_articlenumberRegex	:= '';
_serialnumberRegex	:= '';
_traceID						:= DINT#0;
_activeCheckFQDN		:= FALSE;
_allowedFQDN				:= '';

_previousProcesses.Clear();
END_METHOD

METHOD PUBLIC CopyFrom : BOOL
VAR_INPUT
	IN	: KOSTAL_AF2024_Core_System.I_Interface;
END_VAR

VAR
	_IN		: I_T_ProcessConfig;
//	_udi	: UDINT;
//	_p		: POINTER TO T_PreviousProcess;
//	_resp	: KOSTAL_AF2024_Core_functionResponse.T_functionResponse;
END_VAR

IF NOT SUPER^.CopyFrom(IN) 												THEN RETURN;	END_IF
IF NOT __QUERYINTERFACE(IN, _IN) OR_ELSE _IN = 0 	THEN RETURN;	END_IF

_serialnumberRegex	:= _IN.serialnumberRegex;
_articlenumberRegex	:= _IN.articlenumberRegex;
_traceId						:= _IN.traceId;
_activeCheckFQDN		:= _IN.activeCheckFQDN;
_allowedFQDN				:= _IN.allowedFQDN;

_previousProcesses.CopyFrom(_IN.PreviousProcesses);

CopyFrom:= TRUE;

//FOR _udi:= 1 TO _IN.PreviousProcesses.NumberOfObjects DO

//	IF NOT _previousProcesses.AddObject() THEN RETURN;	END_IF

//	_p:= 	_previousProcesses.Get_P(_previousProcesses.NumberOfObjects, _resp);

//	IF (NOT _resp.success) OR (_p = 0 ) THEN RETURN;	END_IF
	
//	_p^.CopyFrom(IN.IPreviousProcesses.Get_I(_udi, _resp));
		
//END_FOR
END_METHOD

PROPERTY PUBLIC PreviousProcesses : I_ListOfPreviousProcess
GET

PreviousProcesses:= _previousProcesses;
END_GET
END_PROPERTY

PROPERTY PUBLIC PreviousProcesses_Owner : I_ListOfPreviousProcess_Owner
GET

PreviousProcesses_Owner := _previousProcesses;
END_GET
END_PROPERTY

PROPERTY PUBLIC serialnumberRegex : KOSTAL_AF2024_Core_Settings.T_MaxString_UTF8
GET

serialnumberRegex:= _serialnumberRegex;
END_GET
SET

_serialnumberRegex:= serialnumberRegex;
END_SET
END_PROPERTY

PROPERTY PUBLIC traceID : DINT
GET

traceID:= _traceID;
END_GET
SET

_traceID:= traceID;
END_SET
END_PROPERTY

END_FUNCTION_BLOCK

// 3_DUT/SingleProcess/ListOf/FB_ListOfSingleProcess
FUNCTION_BLOCK FB_ListOfSingleProcess  EXTENDS KOSTAL_AF2024_Core_ListOf._FB_Object_Base IMPLEMENTS I_ListOfSingleProcess, I_ListOfSingleProcess_CopyFrom, I_ListOfSingleProcess_Owner

VAR
	_Dummy	: T_SingleProcess;
END_VAR

(*
	Returns the typed interface in the reference variable.
	In the event of an error, the return value becomes FALSE and the interface refers to the {_Dummy}.
*)
METHOD PROTECTED _get_I : I_T_SingleProcess

VAR_INPUT
	Member		: KOSTAL_AF2024_Core_System.I_Interface;
	rValid		: REFERENCE TO BOOL;
	Response	: KOSTAL_AF2024_Core_functionResponse.I_T_functionResponse_Owner;
END_VAR

VAR
	_iObj			: I_T_SingleProcess;
END_VAR
//preset
_get_I:= _Dummy;
IF __ISVALIDREF(rValid)	THEN	rValid:= FALSE;	END_IF	

IF NOT _verifyMember(Member, Response)	THEN RETURN;	END_IF

//return dummy if no valid DUT is found
IF NOT __QUERYINTERFACE(Member, _iObj) OR_ELSE (_iObj = 0)	THEN		
	_setResultFail(Response, "__QueryInterface failed - return Dummy");	RETURN;	
END_IF

IF __ISVALIDREF(rValid)	THEN	rValid:= TRUE;	END_IF	
_setResultPass(Response, "Successful");

_get_I:= _iObj;
END_METHOD

(*
	Returns the typed owner interface in the reference variable.
	In the event of an error, the return value becomes FALSE and the interface refers to the {_Dummy}.
*)
METHOD PROTECTED _get_I_Owner : I_T_SingleProcess_Owner

VAR_INPUT
	Member		: KOSTAL_AF2024_Core_System.I_Interface;
	rValid		: REFERENCE TO BOOL;
	Response	: KOSTAL_AF2024_Core_functionResponse.I_T_functionResponse_Owner;
END_VAR

VAR
	_iObj			: I_T_SingleProcess_Owner;
END_VAR
//preset
_get_I_Owner:= _Dummy;

IF 		__ISVALIDREF(rValid)	THEN	rValid:= FALSE;	END_IF	

IF NOT _verifyMember(Member, Response)	THEN RETURN;	END_IF

//return dummy if no valid DUT is found
IF NOT __QUERYINTERFACE(Member, _iObj) OR_ELSE (_iObj = 0)	THEN	
	_setResultFail(Response, "__QueryInterface failed - return Dummy");	RETURN;	
END_IF

IF __ISVALIDREF(rValid)	THEN	rValid:= TRUE;	END_IF
_setResultPass(Response, "Successful");
_get_I_Owner:= _iObj;
END_METHOD

(*
	Cleans the custom class {FB_DUT} and removes it from memory.
*)
METHOD PROTECTED  _removePayLoad : BOOL
VAR_INPUT
	Member	: KOSTAL_AF2024_Core_System.I_Interface;
	Result	: KOSTAL_AF2024_Core_functionResponse.I_T_functionResponse_Owner;
END_VAR

VAR
	_iObj			: I_T_SingleProcess_Owner;
	_pFB_DUT	:	POINTER TO T_SingleProcess;
	_Success	: BOOL;
END_VAR


IF NOT SUPER^._removePayload(Member, Result)	THEN RETURN;	END_IF

_Success:= __QUERYINTERFACE(Member, _iObj);

IF NOT _Success	THEN	RETURN;	END_IF
IF _iObj = 0		THEN	RETURN;	END_IF

_iObj.Clear();

_Success  := __QUERYPOINTER(_iObj, _pFB_DUT);

IF NOT _Success	THEN	RETURN;	END_IF
IF _pFB_DUT = 0	THEN	RETURN;	END_IF

__DELETE(_pFB_DUT);
END_METHOD

(*
	Overload the method from the base class to verify the custom interface. 
	The local method {_get_I_Owner()} is used for this.
*)
METHOD PROTECTED _verifyMember : BOOL

VAR_INPUT
	Member	: KOSTAL_AF2024_Core_System.I_Interface;
	Result	: KOSTAL_AF2024_Core_functionResponse.I_T_functionResponse_Owner;
END_VAR

VAR
	_pObj	: POINTER TO T_SingleProcess;
	_Success: BOOL;
END_VAR

IF NOT SUPER^._verifyMember(Member, Result)	THEN RETURN;	END_IF

_Success:= __QUERYPOINTER(Member, _pObj);

//return dummy if no valid Pointer to DUT is found
IF NOT _Success OR_ELSE (_pObj = 0)	THEN	_setResultFail(Result, "__QueryPointer failed");	RETURN; END_IF

_verifyMember:= TRUE;
END_METHOD

(*
	Add a new instance of FB_Dut and copy content from [IN] to the new instance
*)
METHOD PUBLIC Add_DUT : BOOL
VAR_INPUT
	IN				: KOSTAL_AF2024_Core_System.I_Interface;
	Response	: KOSTAL_AF2024_Core_functionResponse.I_T_functionResponse_Owner;
END_VAR

VAR
	_IN1	: I_T_SingleProcess;
	_IN2	: I_T_SingleProcess_Owner;
	_pDUT	: POINTER TO T_SingleProcess;
END_VAR

IF IN = 0 THEN	RETURN;	END_IF


IF __QUERYINTERFACE(IN, _IN1) AND_THEN (_IN1 <> 0)	THEN


	_pDUT:= __NEW(T_SingleProcess);
	
	IF _pDUT = 0 THEN	_setResultFail(Response, "cannot create new object"); RETURN; END_IF
	
	_pDUT^.CopyFrom(_IN1);
	
	Add_DUT:= _addMember(_pDUT^, Response);


ELSIF __QUERYINTERFACE(IN, _IN2) AND_THEN (_IN2 <> 0)	THEN


	_pDUT:= __NEW(T_SingleProcess);
	
	IF _pDUT = 0 THEN	_setResultFail(Response, "cannot create new object"); RETURN; END_IF
	
	_pDUT^.CopyFrom(_IN2);
	
	Add_DUT:= _addMember(_pDUT^, Response);


END_IF
END_METHOD

(*
	Makes the protected method public.
*)
METHOD Clear

_clear();
END_METHOD

(*
	Copies the contents of another list {IN} into its own memory.
*)
METHOD PUBLIC CopyFrom
VAR_INPUT
	IN	: KOSTAL_AF2024_Core_System.I_Interface;
END_VAR

VAR
	_udi	: UDINT;

	_IN		: I_ListOfSingleProcess;
	_IN_O	: I_ListOfSingleProcess_Owner;

END_VAR

IF IN = 0 THEN RETURN;	END_IF

IF __QUERYINTERFACE(IN, _IN_O) AND_THEN _IN_O <> 0	THEN

	_clear();
	
	FOR _udi:= 1 TO _IN_O.NumberOfMember DO
		Add_DUT(_IN_O.Get_I_Owner(_udi, 0, 0), 0);
	END_FOR
	
ELSIF __QUERYINTERFACE(IN, _IN) AND_THEN _IN <> 0	THEN	

	_clear();
	
	FOR _udi:= 1 TO _IN.NumberOfMember DO
		Add_DUT(_IN.Get_I(_udi, 0, 0), 0);
	END_FOR

END_IF
END_METHOD

(*
	Copies the own content into another list created at the parameter {IN}.
*)
METHOD PUBLIC CopyTo
VAR_INPUT
	IN	: KOSTAL_AF2024_Core_System.I_Interface;
END_VAR

VAR
	_IN	: I_ListOfSingleProcess_CopyFrom;
END_VAR

IF (IN = 0) OR_ELSE NOT __QUERYINTERFACE(IN, _IN) OR_ELSE (_IN = 0) THEN	RETURN;	END_IF

_IN.CopyFrom(THIS^);
END_METHOD

(*
	Deletes the class specified with the {Number} from the list.
*)
METHOD PUBLIC Delete_DUT : BOOL
VAR_INPUT
	Number		: UDINT;	//Number of DUT in List
	Response	: KOSTAL_AF2024_Core_functionResponse.I_T_functionResponse_Owner;
END_VAR

VAR
	//_response	: KOSTAL_AF2024_Core_functionResponse.T_functionResponse;
	_Success	: BOOL;
	_Member		: KOSTAL_AF2024_Core_System.I_Interface;
END_VAR

IF Number = 0 THEN	_setResultFail(Response, "Number is out of range (1..n)"); RETURN; END_IF

Delete_DUT:= _removeMemberByIndex(Number - 1, Response);
END_METHOD

(*
	Get readonly access to content of Member with {Number}
*) 
METHOD Get_I : I_T_SingleProcess

VAR_INPUT
	Number		: UDINT;
	rValid		: REFERENCE TO BOOL;
	Response	: KOSTAL_AF2024_Core_functionResponse.I_T_functionResponse_Owner;
END_VAR

VAR
	_Member	: KOSTAL_AF2024_Core_System.I_Interface;
END_VAR

//preset
Get_I:=	_Dummy; 
IF __ISVALIDREF(rValid)	THEN	rValid:= FALSE;	END_IF	

IF Number = 0 THEN _setResultFail(Response, "Number is out of range (1..n)"); RETURN; END_IF

IF _findMemberByIndex(Number - 1, _Member, Response) THEN
	Get_I:= _get_I(_Member, rValid, Response);
END_IF
END_METHOD

(*
	Get full access to content of Member with {Number}
*) 
METHOD Get_I_Owner : I_T_SingleProcess_Owner

VAR_INPUT
	Number		: UDINT;
	rValid		: REFERENCE TO BOOL;
	Response	: KOSTAL_AF2024_Core_functionResponse.I_T_functionResponse_Owner;
END_VAR

VAR
	_Member	: KOSTAL_AF2024_Core_System.I_Interface;
END_VAR
//preset

Get_I_Owner:= _Dummy;

IF __ISVALIDREF(rValid)	THEN	rValid:= FALSE;	END_IF	

IF Number = 0 THEN _setResultFail(Response, "Number is out of range (1..n)"); RETURN; END_IF

IF _findMemberByIndex(Number - 1, _Member, Response) THEN
	Get_I_Owner:= _get_I_Owner(_Member, rValid, Response);
END_IF
END_METHOD

(*
	Number of Member in list.
*)
PROPERTY NumberOfMember : UDINT
GET

NumberOfMember:= SUPER^._NumberOfMember;
END_GET
END_PROPERTY

END_FUNCTION_BLOCK

// 3_DUT/SingleProcess/ListOf/I_ListOfSingleProcess
INTERFACE I_ListOfSingleProcess EXTENDS KOSTAL_AF2024_Core_ListOf._I_Object_Base

(*
	Copies the own content into another list created at the parameter {IN}.
*)
METHOD PUBLIC CopyTo
VAR_INPUT
	IN	: KOSTAL_AF2024_Core_System.I_Interface;
END_VAR
END_METHOD

(*
	Get readonly access to content of Member with {Number}
*) 
METHOD Get_I : I_T_SingleProcess

VAR_INPUT
	Number		: UDINT;
	rValid		: REFERENCE TO BOOL;
	Response	: KOSTAL_AF2024_Core_functionResponse.I_T_functionResponse_Owner;
END_VAR
END_METHOD

(*
	Number of Member in list.
*)
PROPERTY NumberOfMember : UDINT
GET
END_GET
END_PROPERTY

END_INTERFACE

// 3_DUT/SingleProcess/I_T_SingleProcess
INTERFACE I_T_SingleProcess EXTENDS _I_T_Copy

PROPERTY PUBLIC articleNumber : KOSTAL_AF2024_Core_Settings.T_MaxString_UTF8
GET
END_GET
END_PROPERTY

PROPERTY PUBLIC id : ULINT
GET
END_GET
END_PROPERTY

PROPERTY PUBLIC OptionalFlags : I_T_OptionalFlags
GET
END_GET
END_PROPERTY

PROPERTY PUBLIC OptionalStrings : I_T_OptionalStrings
GET
END_GET
END_PROPERTY

PROPERTY PUBLIC process : KOSTAL_AF2024_Core_Settings.T_MaxString_UTF8
GET
END_GET
END_PROPERTY

PROPERTY PUBLIC result : BOOL
GET
END_GET
END_PROPERTY

PROPERTY PUBLIC serialNumber : KOSTAL_AF2024_Core_Settings.T_MaxString_UTF8
GET
END_GET
END_PROPERTY

PROPERTY PUBLIC timeStamp : KOSTAL_AF2024_Core_Settings.T_MaxString_UTF8
GET
END_GET
END_PROPERTY

PROPERTY PUBLIC traceId : DINT
GET
END_GET
END_PROPERTY

END_INTERFACE

// 3_DUT/SingleProcess/ListOf/I_ListOfSingleProcess_CopyFrom
INTERFACE I_ListOfSingleProcess_CopyFrom EXTENDS KOSTAL_AF2024_Core_System.I_Interface

METHOD PUBLIC CopyFrom
VAR_INPUT
	IN	: KOSTAL_AF2024_Core_System.I_Interface;
END_VAR
END_METHOD

END_INTERFACE

// 3_DUT/SingleProcess/ListOf/I_ListOfSingleProcess_Owner
INTERFACE I_ListOfSingleProcess_Owner EXTENDS KOSTAL_AF2024_Core_ListOf._I_Object_Base_Owner

(*
	Add a new instance of FB_Dut and copy content from [IN] to the new instance
*)
METHOD PUBLIC Add_DUT : BOOL
VAR_INPUT
	IN				: KOSTAL_AF2024_Core_System.I_Interface;
	Response	: KOSTAL_AF2024_Core_functionResponse.I_T_functionResponse_Owner;
END_VAR
END_METHOD

(*
	Makes the protected method public.
*)
METHOD Clear
END_METHOD

(*
	Copies the contents of another list {IN} into its own memory.
*)
METHOD PUBLIC CopyFrom
VAR_INPUT
	IN	: KOSTAL_AF2024_Core_System.I_Interface;
END_VAR
END_METHOD

(*
	Copies the own content into another list created at the parameter {IN}.
*)
METHOD PUBLIC CopyTo
VAR_INPUT
	IN	: KOSTAL_AF2024_Core_System.I_Interface;
END_VAR
END_METHOD

(*
	Deletes the class specified with the {Number} from the list.
*)
METHOD PUBLIC Delete_DUT : BOOL
VAR_INPUT
	Number		: UDINT;	//Number of DUT in List
	Response	: KOSTAL_AF2024_Core_functionResponse.I_T_functionResponse_Owner;
END_VAR
END_METHOD

(*
	Get readonly access to content of Member with {Number}
*) 
METHOD Get_I : I_T_SingleProcess

VAR_INPUT
	Number		: UDINT;
	rValid		: REFERENCE TO BOOL;
	Response	: KOSTAL_AF2024_Core_functionResponse.I_T_functionResponse_Owner;
END_VAR
END_METHOD

(*
	Get full access to content of Member with {Number}
*) 
METHOD Get_I_Owner : I_T_SingleProcess_Owner

VAR_INPUT
	Number		: UDINT;
	rValid		: REFERENCE TO BOOL;
	Response	: KOSTAL_AF2024_Core_functionResponse.I_T_functionResponse_Owner;
END_VAR
END_METHOD

(*
	Number of Member in list.
*)
PROPERTY NumberOfMember : UDINT
GET
END_GET
END_PROPERTY

END_INTERFACE

// 3_DUT/SingleProcess/I_T_SingleProcess_Owner
INTERFACE I_T_SingleProcess_Owner EXTENDS _I_T_Copy_Owner

PROPERTY PUBLIC articleNumber : KOSTAL_AF2024_Core_Settings.T_MaxString_UTF8
GET
END_GET
SET
END_SET
END_PROPERTY

METHOD PUBLIC clear
VAR_INPUT
END_VAR
END_METHOD

PROPERTY PUBLIC id : ULINT
GET
END_GET
SET
END_SET
END_PROPERTY

PROPERTY PUBLIC OptionalFlags_Owner : I_T_OptionalFlags_Owner
GET
END_GET
END_PROPERTY

PROPERTY PUBLIC OptionalStrings_Owner : I_T_OptionalStrings_Owner
GET
END_GET
END_PROPERTY

PROPERTY PUBLIC process : KOSTAL_AF2024_Core_Settings.T_MaxString_UTF8
GET
END_GET
SET
END_SET
END_PROPERTY

PROPERTY PUBLIC result : BOOL
GET
END_GET
SET
END_SET
END_PROPERTY

PROPERTY PUBLIC serialNumber : KOSTAL_AF2024_Core_Settings.T_MaxString_UTF8
GET
END_GET
SET
END_SET
END_PROPERTY

PROPERTY PUBLIC timeStamp : KOSTAL_AF2024_Core_Settings.T_MaxString_UTF8
GET
END_GET
SET
END_SET
END_PROPERTY

PROPERTY PUBLIC traceId : DINT
GET
END_GET
SET
END_SET
END_PROPERTY

END_INTERFACE

// 3_DUT/SingleProcess/T_SingleProcess
{attribute 'enable_dynamic_creation'}
FUNCTION_BLOCK T_SingleProcess EXTENDS _T_Copy IMPLEMENTS I_T_SingleProcess_Owner, I_T_SingleProcess

VAR
	_id								: ULINT;	//bigint(20)
	_serialNumber			:	KOSTAL_AF2024_Core_Settings.T_MaxString_UTF8;	//varchar(30)
	_articleNumber		:	KOSTAL_AF2024_Core_Settings.T_MaxString_UTF8;	//varchar(30)
	_timeStamp				:	KOSTAL_AF2024_Core_Settings.T_MaxString_UTF8;	//varchar(20)
	_traceId					: DINT;	//int(5)
	_process					:	KOSTAL_AF2024_Core_Settings.T_MaxString_UTF8;		//varchar(10)
	_result						: BOOL;	//tinyint(1)

	_optionalStrings	:	T_OptionalStrings;
	_optionalFlags		: T_OptionalFlags;
END_VAR

PROPERTY PUBLIC articleNumber : KOSTAL_AF2024_Core_Settings.T_MaxString_UTF8
GET

articleNumber:= _articleNumber;
END_GET
SET

_articleNumber:= articleNumber;
END_SET
END_PROPERTY

METHOD PUBLIC clear
VAR_INPUT
END_VAR

_id:= 0;
_serialNumber	:= '';
_articleNumber	:= '';
_timeStamp			:= '';
_traceId				:= 0;
_process				:= '';
_result					:= FALSE;

_optionalStrings.clear();
_optionalFlags.clear();
END_METHOD

METHOD PUBLIC CopyFrom :BOOL
VAR_INPUT
	IN	: KOSTAL_AF2024_Core_System.I_Interface;
END_VAR

VAR
	_IN		: I_T_SingleProcess;
	_IN2	: I_T_SingleProcess_Owner;
END_VAR

IF NOT SUPER^.CopyFrom(IN) THEN RETURN;	END_IF

IF __QUERYINTERFACE(IN, _IN2) AND_THEN _IN2 <> 0 THEN 

	_id						:= _IN2.id;
	_serialNumber	:= _IN2.serialNumber;
	_articleNumber:= _IN2.articleNumber;
	_timeStamp		:= _IN2.timeStamp;
	_traceId			:= _IN2.traceId;
	_process			:= _IN2.process;
	_result				:= _IN2.result;
	
	_optionalStrings.CopyFrom(_IN2.OptionalStrings_Owner);
	_optionalFlags.CopyFrom(_IN2.OptionalFlags_Owner);
	
	CopyFrom:= TRUE;
	
ELSIF __QUERYINTERFACE(IN, _IN) AND_THEN _IN <> 0 THEN 

	_id						:= _IN.id;
	_serialNumber	:= _IN.serialNumber;
	_articleNumber:= _IN.articleNumber;
	_timeStamp		:= _IN.timeStamp;
	_traceId			:= _IN.traceId;
	_process			:= _IN.process;
	_result				:= _IN.result;
	
	_optionalStrings.CopyFrom(_IN.OptionalStrings);
	_optionalFlags.CopyFrom(_IN.OptionalFlags);

	CopyFrom:= TRUE;

END_IF
END_METHOD

PROPERTY PUBLIC id : ULINT
GET

id:= _id;
END_GET
SET

_id:= id;
END_SET
END_PROPERTY

PROPERTY PUBLIC OptionalFlags : I_T_OptionalFlags
GET

OptionalFlags:= _optionalFlags;
END_GET
END_PROPERTY

PROPERTY PUBLIC OptionalFlags_Owner : I_T_OptionalFlags_Owner
GET

OptionalFlags_Owner := _optionalFlags;
END_GET
END_PROPERTY

PROPERTY PUBLIC OptionalStrings : I_T_OptionalStrings
GET

OptionalStrings:= _optionalStrings;
END_GET
END_PROPERTY

PROPERTY PUBLIC OptionalStrings_Owner : I_T_OptionalStrings_Owner
GET

OptionalStrings_Owner := _optionalStrings;
END_GET
END_PROPERTY

PROPERTY PUBLIC process : KOSTAL_AF2024_Core_Settings.T_MaxString_UTF8
GET

process:= _process;
END_GET
SET

_process:= process;
END_SET
END_PROPERTY

PROPERTY PUBLIC result : BOOL
GET

result:= _result;
END_GET
SET

_result:= result;
END_SET
END_PROPERTY

PROPERTY PUBLIC serialNumber : KOSTAL_AF2024_Core_Settings.T_MaxString_UTF8
GET

serialNumber:= _serialNumber;
END_GET
SET

_serialNumber:= serialNumber;
END_SET
END_PROPERTY

PROPERTY PUBLIC timeStamp : KOSTAL_AF2024_Core_Settings.T_MaxString_UTF8
GET

timeStamp:= _timeStamp;
END_GET
SET

_timeStamp:= timeStamp;
END_SET
END_PROPERTY

PROPERTY PUBLIC traceId : DINT
GET

traceId:= _traceId;
END_GET
SET

_traceId:= traceId;
END_SET
END_PROPERTY

END_FUNCTION_BLOCK

// 3_DUT/SubModule/ListOf/FB_ListOfSubModule
FUNCTION_BLOCK FB_ListOfSubModule  EXTENDS KOSTAL_AF2024_Core_ListOf._FB_Object_Base IMPLEMENTS I_ListOfSubModule, I_ListOfSubModule_CopyFrom, I_ListOfSubModule_Owner

VAR
	_Dummy	: T_SubModule;
END_VAR

(*
	Returns the typed interface in the reference variable.
	In the event of an error, the return value becomes FALSE and the interface refers to the {_Dummy}.
*)
METHOD PROTECTED _get_I : I_T_SubModule

VAR_INPUT
	Member		: KOSTAL_AF2024_Core_System.I_Interface;
	rValid		: REFERENCE TO BOOL;
	Response	: KOSTAL_AF2024_Core_functionResponse.I_T_functionResponse_Owner;
END_VAR

VAR
	_iObj			: I_T_SubModule;
END_VAR
//preset
_get_I:= _Dummy;
IF __ISVALIDREF(rValid)	THEN	rValid:= FALSE;	END_IF	

IF NOT _verifyMember(Member, Response)	THEN RETURN;	END_IF

//return dummy if no valid DUT is found
IF NOT __QUERYINTERFACE(Member, _iObj) OR_ELSE (_iObj = 0)	THEN		
	_setResultFail(Response, "__QueryInterface failed - return Dummy");	RETURN;	
END_IF

IF __ISVALIDREF(rValid)	THEN	rValid:= TRUE;	END_IF	
_setResultPass(Response, "Successful");

_get_I:= _iObj;
END_METHOD

(*
	Returns the typed owner interface in the reference variable.
	In the event of an error, the return value becomes FALSE and the interface refers to the {_Dummy}.
*)
METHOD PROTECTED _get_I_Owner : I_T_SubModule_Owner

VAR_INPUT
	Member		: KOSTAL_AF2024_Core_System.I_Interface;
	rValid		: REFERENCE TO BOOL;
	Response	: KOSTAL_AF2024_Core_functionResponse.I_T_functionResponse_Owner;
END_VAR

VAR
	_iObj			: I_T_SubModule_Owner;
END_VAR
//preset
_get_I_Owner:= _Dummy;

IF 		__ISVALIDREF(rValid)	THEN	rValid:= FALSE;	END_IF	

IF NOT _verifyMember(Member, Response)	THEN RETURN;	END_IF

//return dummy if no valid DUT is found
IF NOT __QUERYINTERFACE(Member, _iObj) OR_ELSE (_iObj = 0)	THEN	
	_setResultFail(Response, "__QueryInterface failed - return Dummy");	RETURN;	
END_IF

IF __ISVALIDREF(rValid)	THEN	rValid:= TRUE;	END_IF
_setResultPass(Response, "Successful");
_get_I_Owner:= _iObj;
END_METHOD

(*
	Cleans the custom class {FB_DUT} and removes it from memory.
*)
METHOD PROTECTED  _removePayLoad : BOOL
VAR_INPUT
	Member	: KOSTAL_AF2024_Core_System.I_Interface;
	Result	: KOSTAL_AF2024_Core_functionResponse.I_T_functionResponse_Owner;
END_VAR

VAR
	_iObj			: I_T_SubModule_Owner;
	_pFB_DUT	:	POINTER TO T_SubModule;
	_Success	: BOOL;
END_VAR


IF NOT SUPER^._removePayload(Member, Result)	THEN RETURN;	END_IF

_Success:= __QUERYINTERFACE(Member, _iObj);

IF NOT _Success	THEN	RETURN;	END_IF
IF _iObj = 0		THEN	RETURN;	END_IF

_iObj.Clear();

_Success  := __QUERYPOINTER(_iObj, _pFB_DUT);

IF NOT _Success	THEN	RETURN;	END_IF
IF _pFB_DUT = 0	THEN	RETURN;	END_IF

__DELETE(_pFB_DUT);
END_METHOD

(*
	Overload the method from the base class to verify the custom interface. 
	The local method {_get_I_Owner()} is used for this.
*)
METHOD PROTECTED _verifyMember : BOOL

VAR_INPUT
	Member	: KOSTAL_AF2024_Core_System.I_Interface;
	Result	: KOSTAL_AF2024_Core_functionResponse.I_T_functionResponse_Owner;
END_VAR

VAR
	_pObj	: POINTER TO T_SubModule;
	_Success: BOOL;
END_VAR

IF NOT SUPER^._verifyMember(Member, Result)	THEN RETURN;	END_IF

_Success:= __QUERYPOINTER(Member, _pObj);

//return dummy if no valid Pointer to DUT is found
IF NOT _Success OR_ELSE (_pObj = 0)	THEN	_setResultFail(Result, "__QueryPointer failed");	RETURN; END_IF

_verifyMember:= TRUE;
END_METHOD

(*
	Add a new instance of FB_Dut and copy content from [IN] to the new instance
*)
METHOD PUBLIC Add_DUT : BOOL
VAR_INPUT
	IN				: KOSTAL_AF2024_Core_System.I_Interface;
	Response	: KOSTAL_AF2024_Core_functionResponse.I_T_functionResponse_Owner;
END_VAR

VAR
	_IN1	: I_T_SubModule;
	_IN2	: I_T_SubModule_Owner;
	_pDUT	: POINTER TO T_SubModule;
END_VAR

IF IN = 0 THEN	RETURN;	END_IF


IF __QUERYINTERFACE(IN, _IN1) AND_THEN (_IN1 <> 0)	THEN


	_pDUT:= __NEW(T_SubModule);
	
	IF _pDUT = 0 THEN	_setResultFail(Response, "cannot create new object"); RETURN; END_IF
	
	_pDUT^.CopyFrom(_IN1);
	
	Add_DUT:= _addMember(_pDUT^, Response);


ELSIF __QUERYINTERFACE(IN, _IN2) AND_THEN (_IN2 <> 0)	THEN


	_pDUT:= __NEW(T_SubModule);
	
	IF _pDUT = 0 THEN	_setResultFail(Response, "cannot create new object"); RETURN; END_IF
	
	_pDUT^.CopyFrom(_IN2);
	
	Add_DUT:= _addMember(_pDUT^, Response);


END_IF
END_METHOD

(*
	Makes the protected method public.
*)
METHOD Clear

_clear();
END_METHOD

(*
	Copies the contents of another list {IN} into its own memory.
*)
METHOD PUBLIC CopyFrom
VAR_INPUT
	IN	: KOSTAL_AF2024_Core_System.I_Interface;
END_VAR

VAR
	_udi	: UDINT;

	_IN		: I_ListOfSubModule;
	_IN_O	: I_ListOfSubModule_Owner;

END_VAR

IF IN = 0 THEN RETURN;	END_IF

IF __QUERYINTERFACE(IN, _IN_O) AND_THEN _IN_O <> 0	THEN

	_clear();
	
	FOR _udi:= 1 TO _IN_O.NumberOfMember DO
		Add_DUT(_IN_O.Get_I_Owner(_udi, 0, 0), 0);
	END_FOR
	
ELSIF __QUERYINTERFACE(IN, _IN) AND_THEN _IN <> 0	THEN	

	_clear();
	
	FOR _udi:= 1 TO _IN.NumberOfMember DO
		Add_DUT(_IN.Get_I(_udi, 0, 0), 0);
	END_FOR

END_IF
END_METHOD

(*
	Copies the own content into another list created at the parameter {IN}.
*)
METHOD PUBLIC CopyTo
VAR_INPUT
	IN	: KOSTAL_AF2024_Core_System.I_Interface;
END_VAR

VAR
	_IN	: I_ListOfSubModule_CopyFrom;
END_VAR

IF (IN = 0) OR_ELSE NOT __QUERYINTERFACE(IN, _IN) OR_ELSE (_IN = 0) THEN	RETURN;	END_IF

_IN.CopyFrom(THIS^);
END_METHOD

(*
	Deletes the class specified with the {Number} from the list.
*)
METHOD PUBLIC Delete_DUT : BOOL
VAR_INPUT
	Number		: UDINT;	//Number of DUT in List
	Response	: KOSTAL_AF2024_Core_functionResponse.I_T_functionResponse_Owner;
END_VAR

VAR
	//_response	: KOSTAL_AF2024_Core_functionResponse.T_functionResponse;
	_Success	: BOOL;
	_Member		: KOSTAL_AF2024_Core_System.I_Interface;
END_VAR

IF Number = 0 THEN	_setResultFail(Response, "Number is out of range (1..n)"); RETURN; END_IF

Delete_DUT:= _removeMemberByIndex(Number - 1, Response);
END_METHOD

(*
	Get readonly access to content of Member with {Number}
*) 
METHOD Get_I : I_T_SubModule

VAR_INPUT
	Number		: UDINT;
	rValid		: REFERENCE TO BOOL;
	Response	: KOSTAL_AF2024_Core_functionResponse.I_T_functionResponse_Owner;
END_VAR

VAR
	_Member	: KOSTAL_AF2024_Core_System.I_Interface;
END_VAR

//preset
Get_I:=	_Dummy; 
IF __ISVALIDREF(rValid)	THEN	rValid:= FALSE;	END_IF	

IF Number = 0 THEN _setResultFail(Response, "Number is out of range (1..n)"); RETURN; END_IF

IF _findMemberByIndex(Number - 1, _Member, Response) THEN
	Get_I:= _get_I(_Member, rValid, Response);
END_IF
END_METHOD

(*
	Get full access to content of Member with {Number}
*) 
METHOD Get_I_Owner : I_T_SubModule_Owner

VAR_INPUT
	Number		: UDINT;
	rValid		: REFERENCE TO BOOL;
	Response	: KOSTAL_AF2024_Core_functionResponse.I_T_functionResponse_Owner;
END_VAR

VAR
	_Member	: KOSTAL_AF2024_Core_System.I_Interface;
END_VAR
//preset

Get_I_Owner:= _Dummy;

IF __ISVALIDREF(rValid)	THEN	rValid:= FALSE;	END_IF	

IF Number = 0 THEN _setResultFail(Response, "Number is out of range (1..n)"); RETURN; END_IF

IF _findMemberByIndex(Number - 1, _Member, Response) THEN
	Get_I_Owner:= _get_I_Owner(_Member, rValid, Response);
END_IF
END_METHOD

(*
	Number of Member in list.
*)
PROPERTY NumberOfMember : UDINT
GET

NumberOfMember:= SUPER^._NumberOfMember;
END_GET
END_PROPERTY

END_FUNCTION_BLOCK

// 3_DUT/SubModule/ListOf/I_ListOfSubModule
INTERFACE I_ListOfSubModule EXTENDS KOSTAL_AF2024_Core_ListOf._I_Object_Base

(*
	Copies the own content into another list created at the parameter {IN}.
*)
METHOD PUBLIC CopyTo
VAR_INPUT
	IN	: KOSTAL_AF2024_Core_System.I_Interface;
END_VAR
END_METHOD

(*
	Get readonly access to content of Member with {Number}
*) 
METHOD Get_I : I_T_SubModule

VAR_INPUT
	Number		: UDINT;
	rValid		: REFERENCE TO BOOL;
	Response	: KOSTAL_AF2024_Core_functionResponse.I_T_functionResponse_Owner;
END_VAR
END_METHOD

(*
	Number of Member in list.
*)
PROPERTY NumberOfMember : UDINT
GET
END_GET
END_PROPERTY

END_INTERFACE

// 3_DUT/SubModule/I_T_SubModule
INTERFACE I_T_SubModule EXTENDS _I_T_Copy

PROPERTY PUBLIC articleNumber : KOSTAL_AF2024_Core_Settings.T_MaxString_UTF8
GET
END_GET
END_PROPERTY

PROPERTY PUBLIC serialNumber : KOSTAL_AF2024_Core_Settings.T_MaxString_UTF8
GET
END_GET
END_PROPERTY

END_INTERFACE

// 3_DUT/SubModule/ListOf/I_ListOfSubModule_CopyFrom
INTERFACE I_ListOfSubModule_CopyFrom EXTENDS KOSTAL_AF2024_Core_System.I_Interface

METHOD PUBLIC CopyFrom
VAR_INPUT
	IN	: KOSTAL_AF2024_Core_System.I_Interface;
END_VAR
END_METHOD

END_INTERFACE

// 3_DUT/SubModule/ListOf/I_ListOfSubModule_Owner
INTERFACE I_ListOfSubModule_Owner EXTENDS KOSTAL_AF2024_Core_ListOf._I_Object_Base_Owner

(*
	Add a new instance of FB_Dut and copy content from [IN] to the new instance
*)
METHOD PUBLIC Add_DUT : BOOL
VAR_INPUT
	IN				: KOSTAL_AF2024_Core_System.I_Interface;
	Response	: KOSTAL_AF2024_Core_functionResponse.I_T_functionResponse_Owner;
END_VAR
END_METHOD

(*
	Makes the protected method public.
*)
METHOD Clear
END_METHOD

(*
	Copies the contents of another list {IN} into its own memory.
*)
METHOD PUBLIC CopyFrom
VAR_INPUT
	IN	: KOSTAL_AF2024_Core_System.I_Interface;
END_VAR
END_METHOD

(*
	Copies the own content into another list created at the parameter {IN}.
*)
METHOD PUBLIC CopyTo
VAR_INPUT
	IN	: KOSTAL_AF2024_Core_System.I_Interface;
END_VAR
END_METHOD

(*
	Deletes the class specified with the {Number} from the list.
*)
METHOD PUBLIC Delete_DUT : BOOL
VAR_INPUT
	Number		: UDINT;	//Number of DUT in List
	Response	: KOSTAL_AF2024_Core_functionResponse.I_T_functionResponse_Owner;
END_VAR
END_METHOD

(*
	Get readonly access to content of Member with {Number}
*) 
METHOD Get_I : I_T_SubModule

VAR_INPUT
	Number		: UDINT;
	rValid		: REFERENCE TO BOOL;
	Response	: KOSTAL_AF2024_Core_functionResponse.I_T_functionResponse_Owner;
END_VAR
END_METHOD

(*
	Get full access to content of Member with {Number}
*) 
METHOD Get_I_Owner : I_T_SubModule_Owner

VAR_INPUT
	Number		: UDINT;
	rValid		: REFERENCE TO BOOL;
	Response	: KOSTAL_AF2024_Core_functionResponse.I_T_functionResponse_Owner;
END_VAR
END_METHOD

(*
	Number of Member in list.
*)
PROPERTY NumberOfMember : UDINT
GET
END_GET
END_PROPERTY

END_INTERFACE

// 3_DUT/SubModule/I_T_SubModule_Owner
INTERFACE I_T_SubModule_Owner EXTENDS _I_T_Copy_Owner

PROPERTY PUBLIC articleNumber : KOSTAL_AF2024_Core_Settings.T_MaxString_UTF8
GET
END_GET
SET
END_SET
END_PROPERTY

METHOD PUBLIC clear
END_METHOD

PROPERTY PUBLIC serialNumber : KOSTAL_AF2024_Core_Settings.T_MaxString_UTF8
GET
END_GET
SET
END_SET
END_PROPERTY

END_INTERFACE

// 3_DUT/SubModule/T_SubModule
(*

:Author: Frank Dümpelmann <f.duempelmann@kostal.com>
:Date: 2018-11-02

Function
========
| DATATYPE 
| contains Data set to add a commponent to a part in (SQL) Linecontroller.

Methods and Properties
======================

| PROPERTY PUBLIC serialNumberChild : STRING
| PROPERTY PUBLIC articleNumberChild : STRING

| METHOD PUBLIC clear

*)

{attribute 'enable_dynamic_creation'}
FUNCTION_BLOCK PUBLIC T_SubModule EXTENDS _T_Copy IMPLEMENTS I_T_SubModule_Owner, I_T_SubModule

VAR
	_articleNumber			: KOSTAL_AF2024_Core_Settings.T_MaxString_UTF8;
	_serialNumberChild	: KOSTAL_AF2024_Core_Settings.T_MaxString_UTF8;
END_VAR

PROPERTY PUBLIC articleNumber : KOSTAL_AF2024_Core_Settings.T_MaxString_UTF8
GET

articleNumber:= _articleNumber;
END_GET
SET

_articleNumber:= Tc2_Standard.LEFT(STR:= articleNumber, SIZE:= 30);
END_SET
END_PROPERTY

METHOD PUBLIC clear


_articleNumber		:= '';
_serialNumberChild		:= '';
END_METHOD

METHOD PUBLIC CopyFrom : BOOL
VAR_INPUT
	IN	: KOSTAL_AF2024_Core_System.I_Interface;
END_VAR

VAR
	_IN		: I_T_SubModule;
	_IN2	: I_T_SubModule_Owner;
END_VAR

IF NOT SUPER^.CopyFrom(IN) THEN RETURN;	END_IF

IF __QUERYINTERFACE(IN, _IN2) AND_THEN _IN2 <> 0 THEN 

	_articleNumber		:= _IN2.articleNumber;
	_serialNumberChild:= _IN2.serialNumber;

	CopyFrom:= TRUE;
	
ELSIF __QUERYINTERFACE(IN, _IN) AND_THEN _IN <> 0 THEN 

	_articleNumber		:= _IN.articleNumber;
	_serialNumberChild:= _IN.serialNumber;

	CopyFrom:= TRUE;

END_IF
END_METHOD

PROPERTY PUBLIC serialNumber : KOSTAL_AF2024_Core_Settings.T_MaxString_UTF8
GET

serialNumber:= _serialNumberChild;
END_GET
SET

_serialNumberChild:= Tc2_Standard.LEFT(STR:= serialNumber, SIZE:= 30);
END_SET
END_PROPERTY

END_FUNCTION_BLOCK

// 3_DUT/SubModuleOfProcess/ListOf/FB_ListOfSubModuleOfProcess
FUNCTION_BLOCK FB_ListOfSubModuleOfProcess  EXTENDS KOSTAL_AF2024_Core_ListOf._FB_Object_Base IMPLEMENTS I_ListOfSubModuleOfProcess, I_ListOfSubModuleOfProcess_CopyFrom, I_ListOfSubModuleOfProcess_Owner

VAR
	_Dummy	: T_SubModuleOfProcess;
END_VAR

(*
	Returns the typed interface in the reference variable.
	In the event of an error, the return value becomes FALSE and the interface refers to the {_Dummy}.
*)
METHOD PROTECTED _get_I : I_T_SubModuleOfProcess

VAR_INPUT
	Member		: KOSTAL_AF2024_Core_System.I_Interface;
	rValid		: REFERENCE TO BOOL;
	Response	: KOSTAL_AF2024_Core_functionResponse.I_T_functionResponse_Owner;
END_VAR

VAR
	_iObj			: I_T_SubModuleOfProcess;
END_VAR
//preset
_get_I:= _Dummy;
IF __ISVALIDREF(rValid)	THEN	rValid:= FALSE;	END_IF	

IF NOT _verifyMember(Member, Response)	THEN RETURN;	END_IF

//return dummy if no valid DUT is found
IF NOT __QUERYINTERFACE(Member, _iObj) OR_ELSE (_iObj = 0)	THEN		
	_setResultFail(Response, "__QueryInterface failed - return Dummy");	RETURN;	
END_IF

IF __ISVALIDREF(rValid)	THEN	rValid:= TRUE;	END_IF	
_setResultPass(Response, "Successful");

_get_I:= _iObj;
END_METHOD

(*
	Returns the typed owner interface in the reference variable.
	In the event of an error, the return value becomes FALSE and the interface refers to the {_Dummy}.
*)
METHOD PROTECTED _get_I_Owner : I_T_SubModuleOfProcess_Owner

VAR_INPUT
	Member		: KOSTAL_AF2024_Core_System.I_Interface;
	rValid		: REFERENCE TO BOOL;
	Response	: KOSTAL_AF2024_Core_functionResponse.I_T_functionResponse_Owner;
END_VAR

VAR
	_iObj			: I_T_SubModuleOfProcess_Owner;
END_VAR
//preset
_get_I_Owner:= _Dummy;

IF 		__ISVALIDREF(rValid)	THEN	rValid:= FALSE;	END_IF	

IF NOT _verifyMember(Member, Response)	THEN RETURN;	END_IF

//return dummy if no valid DUT is found
IF NOT __QUERYINTERFACE(Member, _iObj) OR_ELSE (_iObj = 0)	THEN	
	_setResultFail(Response, "__QueryInterface failed - return Dummy");	RETURN;	
END_IF

IF __ISVALIDREF(rValid)	THEN	rValid:= TRUE;	END_IF
_setResultPass(Response, "Successful");
_get_I_Owner:= _iObj;
END_METHOD

(*
	Cleans the custom class {FB_DUT} and removes it from memory.
*)
METHOD PROTECTED  _removePayLoad : BOOL
VAR_INPUT
	Member	: KOSTAL_AF2024_Core_System.I_Interface;
	Result	: KOSTAL_AF2024_Core_functionResponse.I_T_functionResponse_Owner;
END_VAR

VAR
	_iObj			: I_T_SubModuleOfProcess_Owner;
	_pFB_DUT	:	POINTER TO T_SubModuleOfProcess;
	_Success	: BOOL;
END_VAR


IF NOT SUPER^._removePayload(Member, Result)	THEN RETURN;	END_IF

_Success:= __QUERYINTERFACE(Member, _iObj);

IF NOT _Success	THEN	RETURN;	END_IF
IF _iObj = 0		THEN	RETURN;	END_IF

_iObj.Clear();

_Success  := __QUERYPOINTER(_iObj, _pFB_DUT);

IF NOT _Success	THEN	RETURN;	END_IF
IF _pFB_DUT = 0	THEN	RETURN;	END_IF

__DELETE(_pFB_DUT);
END_METHOD

(*
	Overload the method from the base class to verify the custom interface. 
	The local method {_get_I_Owner()} is used for this.
*)
METHOD PROTECTED _verifyMember : BOOL

VAR_INPUT
	Member	: KOSTAL_AF2024_Core_System.I_Interface;
	Result	: KOSTAL_AF2024_Core_functionResponse.I_T_functionResponse_Owner;
END_VAR

VAR
	_pObj	: POINTER TO T_SubModuleOfProcess;
	_Success: BOOL;
END_VAR

IF NOT SUPER^._verifyMember(Member, Result)	THEN RETURN;	END_IF

_Success:= __QUERYPOINTER(Member, _pObj);

//return dummy if no valid Pointer to DUT is found
IF NOT _Success OR_ELSE (_pObj = 0)	THEN	_setResultFail(Result, "__QueryPointer failed");	RETURN; END_IF

_verifyMember:= TRUE;
END_METHOD

(*
	Add a new instance of FB_Dut and copy content from [IN] to the new instance
*)
METHOD PUBLIC Add_DUT : BOOL
VAR_INPUT
	IN				: KOSTAL_AF2024_Core_System.I_Interface;
	Response	: KOSTAL_AF2024_Core_functionResponse.I_T_functionResponse_Owner;
END_VAR

VAR
	_IN1	: I_T_SubModuleOfProcess;
	_IN2	: I_T_SubModuleOfProcess_Owner;
	_pDUT	: POINTER TO T_SubModuleOfProcess;
END_VAR

IF IN = 0 THEN	RETURN;	END_IF


IF __QUERYINTERFACE(IN, _IN1) AND_THEN (_IN1 <> 0)	THEN


	_pDUT:= __NEW(T_SubModuleOfProcess);
	
	IF _pDUT = 0 THEN	_setResultFail(Response, "cannot create new object"); RETURN; END_IF
	
	_pDUT^.CopyFrom(_IN1);
	
	Add_DUT:= _addMember(_pDUT^, Response);


ELSIF __QUERYINTERFACE(IN, _IN2) AND_THEN (_IN2 <> 0)	THEN


	_pDUT:= __NEW(T_SubModuleOfProcess);
	
	IF _pDUT = 0 THEN	_setResultFail(Response, "cannot create new object"); RETURN; END_IF
	
	_pDUT^.CopyFrom(_IN2);
	
	Add_DUT:= _addMember(_pDUT^, Response);


END_IF
END_METHOD

(*
	Makes the protected method public.
*)
METHOD Clear

_clear();
END_METHOD

(*
	Copies the contents of another list {IN} into its own memory.
*)
METHOD PUBLIC CopyFrom
VAR_INPUT
	IN	: KOSTAL_AF2024_Core_System.I_Interface;
END_VAR

VAR
	_udi	: UDINT;

	_IN		: I_ListOfSubModuleOfProcess;
	_IN_O	: I_ListOfSubModuleOfProcess_Owner;

END_VAR

IF IN = 0 THEN RETURN;	END_IF

IF __QUERYINTERFACE(IN, _IN_O) AND_THEN _IN_O <> 0	THEN

	_clear();
	
	FOR _udi:= 1 TO _IN_O.NumberOfMember DO
		Add_DUT(_IN_O.Get_I_Owner(_udi, 0, 0), 0);
	END_FOR
	
ELSIF __QUERYINTERFACE(IN, _IN) AND_THEN _IN <> 0	THEN	

	_clear();
	
	FOR _udi:= 1 TO _IN.NumberOfMember DO
		Add_DUT(_IN.Get_I(_udi, 0, 0), 0);
	END_FOR

END_IF
END_METHOD

(*
	Copies the own content into another list created at the parameter {IN}.
*)
METHOD PUBLIC CopyTo
VAR_INPUT
	IN	: KOSTAL_AF2024_Core_System.I_Interface;
END_VAR

VAR
	_IN	: I_ListOfSubModule_CopyFrom;
END_VAR

IF (IN = 0) OR_ELSE NOT __QUERYINTERFACE(IN, _IN) OR_ELSE (_IN = 0) THEN	RETURN;	END_IF

_IN.CopyFrom(THIS^);
END_METHOD

(*
	Deletes the class specified with the {Number} from the list.
*)
METHOD PUBLIC Delete_DUT : BOOL
VAR_INPUT
	Number		: UDINT;	//Number of DUT in List
	Response	: KOSTAL_AF2024_Core_functionResponse.I_T_functionResponse_Owner;
END_VAR

VAR
	//_response	: KOSTAL_AF2024_Core_functionResponse.T_functionResponse;
	_Success	: BOOL;
	_Member		: KOSTAL_AF2024_Core_System.I_Interface;
END_VAR

IF Number = 0 THEN	_setResultFail(Response, "Number is out of range (1..n)"); RETURN; END_IF

Delete_DUT:= _removeMemberByIndex(Number - 1, Response);
END_METHOD

(*
	Get readonly access to content of Member with {Number}
*) 
METHOD Get_I : I_T_SubModuleOfProcess

VAR_INPUT
	Number		: UDINT;
	rValid		: REFERENCE TO BOOL;
	Response	: KOSTAL_AF2024_Core_functionResponse.I_T_functionResponse_Owner;
END_VAR

VAR
	_Member	: KOSTAL_AF2024_Core_System.I_Interface;
END_VAR

//preset
Get_I:=	_Dummy; 
IF __ISVALIDREF(rValid)	THEN	rValid:= FALSE;	END_IF	

IF Number = 0 THEN _setResultFail(Response, "Number is out of range (1..n)"); RETURN; END_IF

IF _findMemberByIndex(Number - 1, _Member, Response) THEN
	Get_I:= _get_I(_Member, rValid, Response);
END_IF
END_METHOD

(*
	Get full access to content of Member with {Number}
*) 
METHOD Get_I_Owner : I_T_SubModuleOfProcess_Owner

VAR_INPUT
	Number		: UDINT;
	rValid		: REFERENCE TO BOOL;
	Response	: KOSTAL_AF2024_Core_functionResponse.I_T_functionResponse_Owner;
END_VAR

VAR
	_Member	: KOSTAL_AF2024_Core_System.I_Interface;
END_VAR
//preset

Get_I_Owner:= _Dummy;

IF __ISVALIDREF(rValid)	THEN	rValid:= FALSE;	END_IF	

IF Number = 0 THEN _setResultFail(Response, "Number is out of range (1..n)"); RETURN; END_IF

IF _findMemberByIndex(Number - 1, _Member, Response) THEN
	Get_I_Owner:= _get_I_Owner(_Member, rValid, Response);
END_IF
END_METHOD

(*
	Number of Member in list.
*)
PROPERTY NumberOfMember : UDINT
GET

NumberOfMember:= SUPER^._NumberOfMember;
END_GET
END_PROPERTY

END_FUNCTION_BLOCK

// 3_DUT/SubModuleOfProcess/ListOf/I_ListOfSubModuleOfProcess
INTERFACE I_ListOfSubModuleOfProcess EXTENDS KOSTAL_AF2024_Core_ListOf._I_Object_Base

(*
	Copies the own content into another list created at the parameter {IN}.
*)
METHOD PUBLIC CopyTo
VAR_INPUT
	IN	: KOSTAL_AF2024_Core_System.I_Interface;
END_VAR
END_METHOD

(*
	Get readonly access to content of Member with {Number}
*) 
METHOD Get_I : I_T_SubModuleOfProcess

VAR_INPUT
	Number		: UDINT;
	rValid		: REFERENCE TO BOOL;
	Response	: KOSTAL_AF2024_Core_functionResponse.I_T_functionResponse_Owner;
END_VAR
END_METHOD

(*
	Number of Member in list.
*)
PROPERTY NumberOfMember : UDINT
GET
END_GET
END_PROPERTY

END_INTERFACE

// 3_DUT/SubModuleOfProcess/I_T_SubModuleOfProcess
INTERFACE I_T_SubModuleOfProcess EXTENDS I_T_SubModule

PROPERTY PUBLIC timeStamp : KOSTAL_AF2024_Core_Settings.T_MaxString_UTF8
GET
END_GET
END_PROPERTY

END_INTERFACE

// 3_DUT/SubModuleOfProcess/ListOf/I_ListOfSubModuleOfProcess_CopyFrom
INTERFACE I_ListOfSubModuleOfProcess_CopyFrom EXTENDS KOSTAL_AF2024_Core_System.I_Interface

METHOD PUBLIC CopyFrom
VAR_INPUT
	IN	: KOSTAL_AF2024_Core_System.I_Interface;
END_VAR
END_METHOD

END_INTERFACE

// 3_DUT/SubModuleOfProcess/ListOf/I_ListOfSubModuleOfProcess_Owner
INTERFACE I_ListOfSubModuleOfProcess_Owner EXTENDS KOSTAL_AF2024_Core_ListOf._I_Object_Base_Owner

(*
	Add a new instance of FB_Dut and copy content from [IN] to the new instance
*)
METHOD PUBLIC Add_DUT : BOOL
VAR_INPUT
	IN				: KOSTAL_AF2024_Core_System.I_Interface;
	Response	: KOSTAL_AF2024_Core_functionResponse.I_T_functionResponse_Owner;
END_VAR
END_METHOD

(*
	Makes the protected method public.
*)
METHOD Clear
END_METHOD

(*
	Copies the contents of another list {IN} into its own memory.
*)
METHOD PUBLIC CopyFrom
VAR_INPUT
	IN	: KOSTAL_AF2024_Core_System.I_Interface;
END_VAR
END_METHOD

(*
	Copies the own content into another list created at the parameter {IN}.
*)
METHOD PUBLIC CopyTo
VAR_INPUT
	IN	: KOSTAL_AF2024_Core_System.I_Interface;
END_VAR
END_METHOD

(*
	Deletes the class specified with the {Number} from the list.
*)
METHOD PUBLIC Delete_DUT : BOOL
VAR_INPUT
	Number		: UDINT;	//Number of DUT in List
	Response	: KOSTAL_AF2024_Core_functionResponse.I_T_functionResponse_Owner;
END_VAR
END_METHOD

(*
	Get readonly access to content of Member with {Number}
*) 
METHOD Get_I : I_T_SubModuleOfProcess

VAR_INPUT
	Number		: UDINT;
	rValid		: REFERENCE TO BOOL;
	Response	: KOSTAL_AF2024_Core_functionResponse.I_T_functionResponse_Owner;
END_VAR
END_METHOD

(*
	Get full access to content of Member with {Number}
*) 
METHOD Get_I_Owner : I_T_SubModuleOfProcess_Owner

VAR_INPUT
	Number		: UDINT;
	rValid		: REFERENCE TO BOOL;
	Response	: KOSTAL_AF2024_Core_functionResponse.I_T_functionResponse_Owner;
END_VAR
END_METHOD

(*
	Number of Member in list.
*)
PROPERTY NumberOfMember : UDINT
GET
END_GET
END_PROPERTY

END_INTERFACE

// 3_DUT/SubModuleOfProcess/I_T_SubModuleOfProcess_Owner
INTERFACE I_T_SubModuleOfProcess_Owner EXTENDS I_T_SubModule_Owner

PROPERTY PUBLIC timeStamp : KOSTAL_AF2024_Core_Settings.T_MaxString_UTF8
GET
END_GET
SET
END_SET
END_PROPERTY

END_INTERFACE

// 3_DUT/SubModuleOfProcess/T_SubModuleOfProcess
{attribute 'enable_dynamic_creation'}
FUNCTION_BLOCK PUBLIC T_SubModuleOfProcess EXTENDS T_SubModule IMPLEMENTS I_T_SubModuleOfProcess_Owner, I_T_SubModuleOfProcess	//, I_SubModulOfProcess_CopyFrom

VAR
	_timeStamp	: KOSTAL_AF2024_Core_Settings.T_MaxString_UTF8;
END_VAR

METHOD PUBLIC clear

SUPER^.clear();

_timeStamp:= '';
END_METHOD

METHOD PUBLIC CopyFrom : BOOL

VAR_INPUT
	IN	: KOSTAL_AF2024_Core_System.I_Interface;
END_VAR

VAR
	_IN		: I_T_SubModuleOfProcess;
	_IN2	: I_T_SubModuleOfProcess_Owner;

//	_iSubModulOfProcess	: I_T_SubModuleOfProcess;
//	_bResult						: BOOL;
END_VAR

IF NOT SUPER^.CopyFrom(IN) THEN RETURN;	END_IF

IF __QUERYINTERFACE(IN, _IN2) AND_THEN _IN2 <> 0 THEN 

	_timeStamp:= _IN2.timeStamp;
	CopyFrom:= SUPER^.CopyFrom(_IN2);

	
ELSIF __QUERYINTERFACE(IN, _IN) AND_THEN _IN <> 0 THEN 

	_timeStamp:= _IN.timeStamp;
	CopyFrom:= SUPER^.CopyFrom(_IN);

END_IF


//_bResult := __QUERYINTERFACE(IN, _iSubModulOfProcess);

//IF NOT _bResult THEN RETURN;	END_IF
//IF _iSubModulOfProcess = 0 	THEN RETURN;	END_IF

//_timeStamp:= _iSubModulOfProcess.timeStamp;

//SUPER^.CopyFrom(IN);
END_METHOD

PROPERTY PUBLIC timeStamp : KOSTAL_AF2024_Core_Settings.T_MaxString_UTF8
GET

timeStamp:= _timeStamp;
END_GET
SET

_timeStamp:= timeStamp;
END_SET
END_PROPERTY

END_FUNCTION_BLOCK

// 3_DUT/WriteCurrentStampDataDto/I_T_WriteCurrentStampDataDto
INTERFACE I_T_WriteCurrentStampDataDto EXTENDS _I_T_Copy

PROPERTY PUBLIC articleNumber : KOSTAL_AF2024_Core_Settings.T_MaxString_UTF8
GET
END_GET
END_PROPERTY

PROPERTY PUBLIC OptionalFlags : I_T_OptionalFlags
GET
END_GET
END_PROPERTY

PROPERTY PUBLIC OptionalStrings : I_T_OptionalStrings
GET
END_GET
END_PROPERTY

PROPERTY PUBLIC result : BOOL
GET
END_GET
END_PROPERTY

PROPERTY PUBLIC serialNumber : KOSTAL_AF2024_Core_Settings.T_MaxString_UTF8
GET
END_GET
END_PROPERTY

END_INTERFACE

// 3_DUT/WriteCurrentStampDataDto/I_T_WriteCurrentStampDataDto_Owner
INTERFACE I_T_WriteCurrentStampDataDto_Owner EXTENDS _I_T_Copy_Owner

PROPERTY PUBLIC articleNumber : KOSTAL_AF2024_Core_Settings.T_MaxString_UTF8
GET
END_GET
SET
END_SET
END_PROPERTY

METHOD PUBLIC clear
VAR_INPUT
END_VAR
END_METHOD

PROPERTY PUBLIC OptionalFlags_Owner : I_T_OptionalFlags_Owner
GET
END_GET
END_PROPERTY

PROPERTY PUBLIC OptionalStrings_Owner : I_T_OptionalStrings_Owner
GET
END_GET
END_PROPERTY

PROPERTY PUBLIC result : BOOL
GET
END_GET
SET
END_SET
END_PROPERTY

PROPERTY PUBLIC serialNumber : KOSTAL_AF2024_Core_Settings.T_MaxString_UTF8
GET
END_GET
SET
END_SET
END_PROPERTY

END_INTERFACE

// 3_DUT/WriteCurrentStampDataDto/T_WriteCurrentStampDataDto
FUNCTION_BLOCK T_WriteCurrentStampDataDto EXTENDS _T_Copy IMPLEMENTS I_T_WriteCurrentStampDataDto_Owner, I_T_WriteCurrentStampDataDto

VAR
	_serialNumber			:	KOSTAL_AF2024_Core_Settings.T_MaxString_UTF8;	//varchar(30)
	_articleNumber		:	KOSTAL_AF2024_Core_Settings.T_MaxString_UTF8;	//varchar(30)
	_result						: BOOL;	//tinyint(1)

	_optionalStrings	:	T_OptionalStrings;
	_optionalFlags		: T_OptionalFlags;
END_VAR

PROPERTY PUBLIC articleNumber : KOSTAL_AF2024_Core_Settings.T_MaxString_UTF8
GET

articleNumber:= _articleNumber;
END_GET
SET

_articleNumber:= articleNumber;
END_SET
END_PROPERTY

METHOD PUBLIC clear
VAR_INPUT
END_VAR

_serialNumber		:= '';
_articleNumber	:= '';
_result					:= FALSE;

_optionalStrings.clear();
_optionalFlags.clear();
END_METHOD

METHOD PUBLIC CopyFrom : BOOL
VAR_INPUT
	IN	: KOSTAL_AF2024_Core_System.I_Interface;
END_VAR

VAR
	_IN		: I_T_WriteCurrentStampDataDto;
	_IN2	: I_T_WriteCurrentStampDataDto_Owner;
END_VAR

IF NOT SUPER^.CopyFrom(IN) THEN ;	

ELSIF __QUERYINTERFACE(IN, _IN2) AND_THEN _IN2 <> 0 THEN 

	_serialNumber			:= _IN2.serialNumber;
	_articleNumber		:= _IN2.articleNumber;
	_result						:= _IN2.result;
	
	_optionalStrings.CopyFrom(_IN2.OptionalStrings_Owner);
	_optionalFlags.CopyFrom(_IN2.OptionalFlags_Owner);

ELSIF __QUERYINTERFACE(IN, _IN) AND_THEN _IN <> 0 THEN 

	_serialNumber			:= _IN.serialNumber;
	_articleNumber		:= _IN.articleNumber;
	_result						:= _IN.result;
	
	_optionalStrings.CopyFrom(_IN.OptionalStrings);
	_optionalFlags.CopyFrom(_IN.OptionalFlags);

END_IF
END_METHOD

PROPERTY PUBLIC OptionalFlags : I_T_OptionalFlags
GET

OptionalFlags:= _optionalFlags;
END_GET
END_PROPERTY

PROPERTY PUBLIC OptionalFlags_Owner : I_T_OptionalFlags_Owner
GET

OptionalFlags_Owner := _optionalFlags;
END_GET
END_PROPERTY

PROPERTY PUBLIC OptionalStrings : I_T_OptionalStrings
GET

OptionalStrings:= _optionalStrings;
END_GET
END_PROPERTY

PROPERTY PUBLIC OptionalStrings_Owner : I_T_OptionalStrings_Owner
GET

OptionalStrings_Owner := _optionalStrings;
END_GET
END_PROPERTY

PROPERTY PUBLIC result : BOOL
GET

result:= _result;
END_GET
SET

_result:= result;
END_SET
END_PROPERTY

PROPERTY PUBLIC serialNumber : KOSTAL_AF2024_Core_Settings.T_MaxString_UTF8
GET

serialNumber:= _serialNumber;
END_GET
SET

_serialNumber:= serialNumber;
END_SET
END_PROPERTY

END_FUNCTION_BLOCK

// 5_POU/GetetParentBySubmoduleSerialnumber/FB_GetParent_By_SM_SN
(*
|MUST EXEND
|
|Extends the base WebService LC with a 
|read
|and a 
|read previous Stamp 
|functionality
*)
FUNCTION_BLOCK PUBLIC FB_GetParent_By_SM_SN EXTENDS FB_LC

VAR

	//======================================================================================
	//Read
	//======================================================================================
	
	//======================================================================================
	//do not insert to _DELETE() !!!!
	//======================================================================================

	
	//======================================================================================
	//Response
	//======================================================================================

	_ResponseProcess	: T_SingleProcess;

	_JsonProcessInfo			: Tc3_IotBase.SJsonValue;

	_JsonSubModules				: Tc3_IotBase.SJsonValue;
	_SubModuleListLenght	: UDINT;

	_ListOfSubModules	: FB_ListOfSubModuleOfProcess;

	//======================================================================================
	//Parameter
	//======================================================================================
	_SerialNumber			: KOSTAL_AF2024_Core_Settings.T_MaxString_UTF8;

END_VAR

VAR CONSTANT
	_ADDRESS_FINISH_FAIL : INT:= 100;
END_VAR

(*
	| return the Process Info from List with {Index} (Base = 0)
*)
METHOD PROTECTED _getProcessInfo : KOSTAL_AF2024_Core_Settings.T_MaxString_UTF8

VAR_INPUT
	IN		: Tc3_IotBase.SJsonValue;
END_VAR

VAR
	_J	: Tc3_IotBase.SJsonValue;
	_uliResult: ULINT;
	_udiResult: UDINT;
	_diResult	: DINT;
	_bResult	: BOOL;
	_sResult	: KOSTAL_AF2024_Core_Settings.T_MaxString_UTF8;
END_VAR

_ResponseProcess.clear();

IF IN = 0 THEN _getProcessInfo:= 'IN Parameter is empty';	RETURN;	END_IF

_sResp:= _PARSE_JSON(IN, PROCESS_INFO.processInfo, _J);
IF _sResp <> '' THEN	_getProcessInfo:= _sResp;	RETURN; END_IF
IF _J = 0	THEN _getProcessInfo:= '_getProcessInfo - no content availabe';	RETURN;	END_IF

_JsonProcessInfo:= _J;

_sResp:= _PARSE_ULINT(_J, PROCESS_INFO.id, _uliResult);
IF _sResp <> '' THEN	_getProcessInfo:= _sResp;	ELSE	_ResponseProcess.id:= _uliResult; END_IF

_sResp:= _PARSE_STRING(_J, PROCESS_INFO.serialNumber, _sResult);
IF _sResp <> '' THEN	_getProcessInfo:= _sResp;	ELSE	_ResponseProcess.serialNumber:= _sResult;	END_IF

_sResp:= _PARSE_STRING(_J, PROCESS_INFO.articleNumber, _sResult);
IF _sResp <> '' THEN	_getProcessInfo:= _sResp;	ELSE	_ResponseProcess.articleNumber:= _sResult;	END_IF

_sResp:= _PARSE_STRING(_J, PROCESS_INFO.timeStamp, _sResult);
IF _sResp <> '' THEN	_getProcessInfo:= _sResp;	ELSE	_ResponseProcess.timeStamp:= _sResult;	END_IF

_sResp:= _PARSE_DINT(_J, PROCESS_INFO.traceId, _diResult);
IF _sResp <> '' THEN	_getProcessInfo:= _sResp;	ELSE	_ResponseProcess.traceId:= _diResult; END_IF

_sResp:= _PARSE_STRING(_J, PROCESS_INFO.process, _sResult);
IF _sResp <> '' THEN	_getProcessInfo:= _sResp;	ELSE	_ResponseProcess.process:= _sResult;	END_IF

_sResp:= _PARSE_BOOL(_J, PROCESS_INFO.result, _bResult);
IF _sResp <> '' THEN	_getProcessInfo:= _sResp;	ELSE	_ResponseProcess.result:= _bResult;	END_IF

_sResp:= _PARSE_STRING(_J, PROCESS_INFO.optionalString_1, _sResult);
IF _sResp <> '' THEN	_getProcessInfo:= _sResp;	ELSE	_ResponseProcess.OptionalStrings_Owner.set(1, _sResult);	END_IF

_sResp:= _PARSE_STRING(_J, PROCESS_INFO.optionalString_2, _sResult);
IF _sResp <> '' THEN	_getProcessInfo:= _sResp;	ELSE	_ResponseProcess.OptionalStrings_Owner.set(2, _sResult);	END_IF

_sResp:= _PARSE_STRING(_J, PROCESS_INFO.optionalString_3, _sResult);
IF _sResp <> '' THEN	_getProcessInfo:= _sResp;	ELSE	_ResponseProcess.OptionalStrings_Owner.set(3, _sResult);	END_IF

_sResp:= _PARSE_STRING(_J, PROCESS_INFO.optionalString_4, _sResult);
IF _sResp <> '' THEN	_getProcessInfo:= _sResp;	ELSE	_ResponseProcess.OptionalStrings_Owner.set(4, _sResult);	END_IF

_sResp:= _PARSE_BOOL(_J, PROCESS_INFO.optionalFlag_1, _bResult);
IF _sResp <> '' THEN	_getProcessInfo:= _sResp;	ELSE	_ResponseProcess.OptionalFlags_Owner.set(1, (_bResult <> 0));	END_IF

_sResp:= _PARSE_BOOL(_J, PROCESS_INFO.optionalFlag_2, _bResult);
IF _sResp <> '' THEN	_getProcessInfo:= _sResp;	ELSE	_ResponseProcess.OptionalFlags_Owner.set(2, (_bResult <> 0));	END_IF

_sResp:= _PARSE_BOOL(_J, PROCESS_INFO.optionalFlag_3, _bResult);
IF _sResp <> '' THEN	_getProcessInfo:= _sResp;	ELSE	_ResponseProcess.OptionalFlags_Owner.set(3, (_bResult <> 0));	END_IF

_sResp:= _PARSE_BOOL(_J, PROCESS_INFO.optionalFlag_4, _bResult);
IF _sResp <> '' THEN	_getProcessInfo:= _sResp;	ELSE	_ResponseProcess.OptionalFlags_Owner.set(4, (_bResult <> 0));	END_IF

_sResp:= _PARSE_BOOL(_J, PROCESS_INFO.optionalFlag_5, _bResult);
IF _sResp <> '' THEN	_getProcessInfo:= _sResp;	ELSE	_ResponseProcess.OptionalFlags_Owner.set(5, (_bResult <> 0));	END_IF

_sResp:= _PARSE_BOOL(_J, PROCESS_INFO.optionalFlag_6, _bResult);
IF _sResp <> '' THEN	_getProcessInfo:= _sResp;	ELSE	_ResponseProcess.OptionalFlags_Owner.set(6, (_bResult <> 0));	END_IF

_sResp:= _PARSE_BOOL(_J, PROCESS_INFO.optionalFlag_7, _bResult);
IF _sResp <> '' THEN	_getProcessInfo:= _sResp;	ELSE	_ResponseProcess.OptionalFlags_Owner.set(7, (_bResult <> 0));	END_IF

_sResp:= _PARSE_BOOL(_J, PROCESS_INFO.optionalFlag_8, _bResult);
IF _sResp <> '' THEN	_getProcessInfo:= _sResp;	ELSE	_ResponseProcess.OptionalFlags_Owner.set(8, (_bResult <> 0));	END_IF
END_METHOD

METHOD PROTECTED _getSubModule_n : KOSTAL_AF2024_Core_Settings.T_MaxString_UTF8

VAR_INPUT
	IN		: Tc3_IotBase.SJsonValue;
	Index	: UDINT;
END_VAR

VAR
	_IN				: Tc3_IotBase.SJsonValue;
	_J				: Tc3_IotBase.SJsonValue;
	_sResult	: KOSTAL_AF2024_Core_Settings.T_MaxString_UTF8;
	_SP				: T_SubModuleOfProcess;
END_VAR
IF IN = 0 												THEN _getSubModule_n:= 'IN Parameter is empty';												RETURN;	END_IF
//IF Index = 0 										THEN _getSubModule_n:= 'Index is out of Range (Base = 1';							RETURN;	END_IF
IF _SubModuleListLenght = 0				THEN _getSubModule_n:= 'no content available';												RETURN;	END_IF
IF Index >= _SubModuleListLenght	THEN _getSubModule_n:= 'Index is out of Range';												RETURN;	END_IF

_J:= _JsonParser.GetArrayValueByIdx(IN,Index);

IF _J = 0	THEN _getSubModule_n:= '_getSubModule_n - no content availabe';	RETURN;	END_IF

_SP.clear();

_PARSE_STRING(_J, SUBMODUL_INFO.articleNumber, _sResult);	
_SP.articleNumber:= _sResult;

_PARSE_STRING(_J, SUBMODUL_INFO.serialNumber, _sResult);
_SP.serialNumber:= _sResult;

_PARSE_STRING(_J, SUBMODUL_INFO.timestamp, _sResult);
_SP.timeStamp:= _sResult;

_ListOfSubModules.Add_DUT(_SP, 0);



(*
IF IN = 0 THEN _getSubModules:= 'IN Parameter is empty';	RETURN;	END_IF

_sResp:= _PARSE_JSON(IN, PROCESS_INFO.processInfo, _IN);
IF _sResp <> '' THEN	_getSubModules:= _sResp;	RETURN; END_IF

_sResp:= _PARSE_ARRAY(_IN, SUBMODUL_INFO.subModules, _J);
IF _sResp <> '' THEN	_getSubModules:= _sResp;	RETURN; END_IF
IF _J = 0	THEN _getSubModules:= '_getSubModules - no content availabe';	RETURN;	END_IF

_jIterator		:= _JsonParser.ArrayBegin(_J);
_jIteratorEnd	:= _JsonParser.ArrayEnd(_J);

WHILE _jIterator <> _jIteratorEnd DO 
	
  _jElement := _JsonParser.GetArrayValue(_jIterator);
	IF _jElement = 0 THEN _getSubModules:= '_getSubModules - sub module corrupt';	RETURN;	END_IF

	_ListOfSubModules.AddObject();
	_pLoSM:= _ListOfSubModules.Get_P(_ListOfSubModules.NumberOfObjects, 0);
	
	_sResp:= _PARSE_STRING(_J, SUBMODUL_INFO.articleNumber, _sResult);
	IF _sResp <> '' THEN	_getSubModules:= _sResp;	ELSE	_pLoSM^.articleNumber:=_sResult;	END_IF

	_sResp:= _PARSE_STRING(_J, SUBMODUL_INFO.serialNumber, _sResult);
	IF _sResp <> '' THEN	_getSubModules:= _sResp;	ELSE	_pLoSM^.serialNumber:=_sResult;	END_IF

	_sResp:= _PARSE_STRING(_J, SUBMODUL_INFO.timestamp, _sResult);
	IF _sResp <> '' THEN	_getSubModules:= _sResp;	ELSE	_pLoSM^.timeStamp:=_sResult;	END_IF
	
  _jIterator := _JsonParser.NextArray(_jIterator);

END_WHILE


*)
END_METHOD

METHOD PROTECTED _getSubModuleList : KOSTAL_AF2024_Core_Settings.T_MaxString_UTF8
VAR_INPUT
	IN	: Tc3_IotBase.SJsonValue;
END_VAR

IF IN = 0 THEN _getSubModuleList:= '_getSubModuleList - IN Parameter is empty';	RETURN;	END_IF

_SubModuleListLenght:= 0;

_getSubModuleList:= _PARSE_ARRAY(IN, SUBMODUL_INFO.subModules, _JsonSubModules);

IF _getSubModuleList <> '' THEN	RETURN;	END_IF

_SubModuleListLenght:=  _JsonParser.GetArraySize(_JsonSubModules);
END_METHOD

METHOD PROTECTED _01_Ready : BOOL
VAR_INPUT
END_VAR


IF NOT 	SUPER^._01_Ready() 								THEN	

	;

ELSIF		_THIS_CALLED = E_PROCESS.idle			THEN	

	_state.clear();	
	_state.ready:= TRUE;

ELSIF		_THIS_CALLED = E_PROCESS.execute	THEN	

	_THIS_IN_PROCESS:= _THIS_CALLED;	

	_state.clear();	
	_state.busy:= TRUE;

	_selectUrl();

	_step.INC();

ELSE

	_state.clear();
	_state.fail:= TRUE;
	_state.description:= Tc2_Standard.WCONCAT("Unknown Process called:", INT_TO_WSTRING(_THIS_CALLED));
	
END_IF
END_METHOD

METHOD PROTECTED _10_getProcessInfo
VAR_INPUT
END_VAR

IF _step.toggle THEN
	;
END_IF

_sResp:= _getProcessInfo(_jsonDoc);

IF _sResp <> '' THEN
	
	_state.clear();
	_state.description:= Tc2_Standard.WCONCAT("Process Info is corrupt;", TO_WSTRING(_sResp));
	_step.set(_ADDRESS_FINISH_FAIL);

ELSE	

	_step.INC();

END_IF
END_METHOD

METHOD PROTECTED _10_getSubModule_n
VAR_INPUT
END_VAR

IF _step.toggle THEN
	;
END_IF

IF _ListOfSubModules.NumberOfMember < _SubModuleListLenght THEN

	_sResp:= _getSubModule_n(_JsonSubModules,  _ListOfSubModules.NumberOfMember);

	IF _sResp <> '' THEN
		
		_state.clear();
		_state.description:= Tc2_Standard.WCONCAT("Sub Module List is corrupt;", TO_WSTRING(_sResp));
		_step.set(_ADDRESS_FINISH_FAIL);
	
	END_IF

ELSE

	_step.INC();

END_IF


(*

_getSubModules(_JsonSubModules);

_step.INC();


//Sub modules are optional
_sResp:= _getSubModules(_jsonDoc);

IF _sResp <> '' THEN
	
	_state.clear();
	_state.description:= Tc2_Standard.CONCAT('Process Info is corrupt;', _sResp);
	_step.set(_ADDRESS_FINISH_FAIL);

ELSE	

	_step.INC();

END_IF
*)
END_METHOD

METHOD PROTECTED _10_getSubModuleList
VAR_INPUT
END_VAR

IF _step.toggle THEN
	;
END_IF

_sResp:= _getSubModuleList(_JsonProcessInfo);

IF _sResp <> '' THEN

	_state.clear();
	_state.description:= Tc2_Standard.WCONCAT("ProcessListInfo is corrupt;", TO_WSTRING(_sResp));
	
	_step.set(_ADDRESS_FINISH_FAIL);

ELSIF _SubModuleListLenght = 0 THEN
	
	_state.clear();
	_state.description:= "no SubModuleList available";

	_step.set(_ADDRESS_FINISH_FAIL);

ELSE
	
	_step.INC();

END_IF
END_METHOD

METHOD PROTECTED _10_processRead
VAR_INPUT
END_VAR

IF _step.toggle THEN

	_JsonProcessInfo:= 0;
	
	_ResponseResult.clear();
	_ResponseProcess.clear();
	_ListOfSubModules.Clear();

END_IF

_00_clientCfg();
END_METHOD

(*
| MUST EXTEND
*)
METHOD PROTECTED _selectUrl


_sUrl:= _UriGet(URL.READ_PARENT_BY_SUB_MODULE_SERIAL_NUMBER);

_UrlReplace(_sUrl, URL.PLACEHOLDER_CLIENT_NAME, _ClientName);
_UrlReplace(_sUrl, URL.PLACEHOLDER_CLIENT_PROCESS, _ClientProcess);
_UrlReplace(_sUrl, URL.PLACEHOLDER_SUB_MODULE_SERIAL_NUMBER, _SerialNumber);
END_METHOD

(*
*)
METHOD Execute : BOOL

VAR_INPUT
	SerialNumber		: KOSTAL_AF2024_Core_Settings.T_MaxString_UTF8;
END_VAR

IF _THIS_CALLED <> E_PROCESS.idle THEN Execute:= FALSE;	RETURN; END_IF

_THIS_CALLED:= E_PROCESS.execute;

IF NOT MT_Usage THEN _SerialNumber	:= SerialNumber;	END_IF

_FBmain();

Execute:= _THIS_CALLED = _THIS_IN_PROCESS;
END_METHOD

PROPERTY PUBLIC ListOfSubModules : I_ListOfSubModuleOfProcess
GET

ListOfSubModules	:= _ListOfSubModules;
END_GET
END_PROPERTY

PROPERTY PUBLIC ResponseProcess : I_T_SingleProcess
GET

ResponseProcess:= _ResponseProcess;
END_GET
END_PROPERTY

PROPERTY ResponseResult : I_T_ResponseResult
GET

ResponseResult := _ResponseResult;
END_GET
END_PROPERTY

METHOD PROTECTED _FBmain
VAR_INPUT
END_VAR

SUPER^._FBmain();

CASE _step.actual OF

	0:	_01_Ready();
	//
	1:	_10_processRead();
	2:	_10_GET();
	3:	_10_GET_CTRL();
	4:	_10_GET_ResponseResult(TRUE);
	5:	_10_GET_ResponseResult_CTRL();
	6:	_10_getProcessInfo();
	7:	_10_getSubModuleList();
	8:	_10_getSubModule_n();
	9:	_10_finishPass();

	100:	_10_finishFail();
ELSE
	
	_99_stepError();
		
END_CASE
END_METHOD

END_FUNCTION_BLOCK

// 5_POU/GetSubModulesByParentSerialNumber/FB_GetSM_ByParentSN
(*
|MUST EXEND
|
|Extends the base WebService LC with a 
|read
|and a 
|read previous Stamp 
|functionality
*)
FUNCTION_BLOCK PUBLIC FB_GetSM_ByParentSN EXTENDS FB_LC

VAR

	//======================================================================================
	//Read
	//======================================================================================
	
	//======================================================================================
	//do not insert to _DELETE() !!!!
	//======================================================================================

	
	//======================================================================================
	//Response
	//======================================================================================

	_ResponseProcess	: T_SingleProcess;

	_JsonProcessInfo			: Tc3_IotBase.SJsonValue;

	_JsonSubModules				: Tc3_IotBase.SJsonValue;
	_SubModuleListLenght	: UDINT;

	_ListOfSubModules	: FB_ListOfSubModuleOfProcess;

	//======================================================================================
	//Parameter
	//======================================================================================
	_SerialNumber			: KOSTAL_AF2024_Core_Settings.T_MaxString_UTF8;

END_VAR

VAR CONSTANT
	_ADDRESS_FINISH_FAIL : INT:= 100;
END_VAR

(*
	| return the Process Info from List with {Index} (Base = 0)
*)
METHOD PROTECTED _getProcessInfo : KOSTAL_AF2024_Core_Settings.T_MaxString_UTF8

VAR_INPUT
	IN		: Tc3_IotBase.SJsonValue;
END_VAR

VAR
	_J	: Tc3_IotBase.SJsonValue;
	_uliResult: ULINT;
	_udiResult: UDINT;
	_diResult	: DINT;
	_bResult	: BOOL;
	_sResult	: KOSTAL_AF2024_Core_Settings.T_MaxString_UTF8;
END_VAR

_ResponseProcess.clear();

IF IN = 0 THEN _getProcessInfo:= 'IN Parameter is empty';	RETURN;	END_IF

_sResp:= _PARSE_JSON(IN, PROCESS_INFO.processInfo, _J);
IF _sResp <> '' THEN	_getProcessInfo:= _sResp;	RETURN; END_IF
IF _J = 0	THEN _getProcessInfo:= '_getProcessInfo - no content availabe';	RETURN;	END_IF

_JsonProcessInfo:= _J;

_sResp:= _PARSE_ULINT(_J, PROCESS_INFO.id, _uliResult);
IF _sResp <> '' THEN	_getProcessInfo:= _sResp;	ELSE	_ResponseProcess.id:= _uliResult; END_IF

_sResp:= _PARSE_STRING(_J, PROCESS_INFO.serialNumber, _sResult);
IF _sResp <> '' THEN	_getProcessInfo:= _sResp;	ELSE	_ResponseProcess.serialNumber:= _sResult;	END_IF

_sResp:= _PARSE_STRING(_J, PROCESS_INFO.articleNumber, _sResult);
IF _sResp <> '' THEN	_getProcessInfo:= _sResp;	ELSE	_ResponseProcess.articleNumber:= _sResult;	END_IF

_sResp:= _PARSE_STRING(_J, PROCESS_INFO.timeStamp, _sResult);
IF _sResp <> '' THEN	_getProcessInfo:= _sResp;	ELSE	_ResponseProcess.timeStamp:= _sResult;	END_IF

_sResp:= _PARSE_DINT(_J, PROCESS_INFO.traceId, _diResult);
IF _sResp <> '' THEN	_getProcessInfo:= _sResp;	ELSE	_ResponseProcess.traceId:= _diResult; END_IF

_sResp:= _PARSE_STRING(_J, PROCESS_INFO.process, _sResult);
IF _sResp <> '' THEN	_getProcessInfo:= _sResp;	ELSE	_ResponseProcess.process:= _sResult;	END_IF

_sResp:= _PARSE_BOOL(_J, PROCESS_INFO.result, _bResult);
IF _sResp <> '' THEN	_getProcessInfo:= _sResp;	ELSE	_ResponseProcess.result:= _bResult;	END_IF

_sResp:= _PARSE_STRING(_J, PROCESS_INFO.optionalString_1, _sResult);
IF _sResp <> '' THEN	_getProcessInfo:= _sResp;	ELSE	_ResponseProcess.OptionalStrings_Owner.set(1, _sResult);	END_IF

_sResp:= _PARSE_STRING(_J, PROCESS_INFO.optionalString_2, _sResult);
IF _sResp <> '' THEN	_getProcessInfo:= _sResp;	ELSE	_ResponseProcess.OptionalStrings_Owner.set(2, _sResult);	END_IF

_sResp:= _PARSE_STRING(_J, PROCESS_INFO.optionalString_3, _sResult);
IF _sResp <> '' THEN	_getProcessInfo:= _sResp;	ELSE	_ResponseProcess.OptionalStrings_Owner.set(3, _sResult);	END_IF

_sResp:= _PARSE_STRING(_J, PROCESS_INFO.optionalString_4, _sResult);
IF _sResp <> '' THEN	_getProcessInfo:= _sResp;	ELSE	_ResponseProcess.OptionalStrings_Owner.set(4, _sResult);	END_IF

_sResp:= _PARSE_BOOL(_J, PROCESS_INFO.optionalFlag_1, _bResult);
IF _sResp <> '' THEN	_getProcessInfo:= _sResp;	ELSE	_ResponseProcess.OptionalFlags_Owner.set(1, (_bResult <> 0));	END_IF

_sResp:= _PARSE_BOOL(_J, PROCESS_INFO.optionalFlag_2, _bResult);
IF _sResp <> '' THEN	_getProcessInfo:= _sResp;	ELSE	_ResponseProcess.OptionalFlags_Owner.set(2, (_bResult <> 0));	END_IF

_sResp:= _PARSE_BOOL(_J, PROCESS_INFO.optionalFlag_3, _bResult);
IF _sResp <> '' THEN	_getProcessInfo:= _sResp;	ELSE	_ResponseProcess.OptionalFlags_Owner.set(3, (_bResult <> 0));	END_IF

_sResp:= _PARSE_BOOL(_J, PROCESS_INFO.optionalFlag_4, _bResult);
IF _sResp <> '' THEN	_getProcessInfo:= _sResp;	ELSE	_ResponseProcess.OptionalFlags_Owner.set(4, (_bResult <> 0));	END_IF

_sResp:= _PARSE_BOOL(_J, PROCESS_INFO.optionalFlag_5, _bResult);
IF _sResp <> '' THEN	_getProcessInfo:= _sResp;	ELSE	_ResponseProcess.OptionalFlags_Owner.set(5, (_bResult <> 0));	END_IF

_sResp:= _PARSE_BOOL(_J, PROCESS_INFO.optionalFlag_6, _bResult);
IF _sResp <> '' THEN	_getProcessInfo:= _sResp;	ELSE	_ResponseProcess.OptionalFlags_Owner.set(6, (_bResult <> 0));	END_IF

_sResp:= _PARSE_BOOL(_J, PROCESS_INFO.optionalFlag_7, _bResult);
IF _sResp <> '' THEN	_getProcessInfo:= _sResp;	ELSE	_ResponseProcess.OptionalFlags_Owner.set(7, (_bResult <> 0));	END_IF

_sResp:= _PARSE_BOOL(_J, PROCESS_INFO.optionalFlag_8, _bResult);
IF _sResp <> '' THEN	_getProcessInfo:= _sResp;	ELSE	_ResponseProcess.OptionalFlags_Owner.set(8, (_bResult <> 0));	END_IF
END_METHOD

METHOD PROTECTED _getSubModule_n : KOSTAL_AF2024_Core_Settings.T_MaxString_UTF8

VAR_INPUT
	IN		: Tc3_IotBase.SJsonValue;
	Index	: UDINT;
END_VAR

VAR
	_IN				: Tc3_IotBase.SJsonValue;
	_J				: Tc3_IotBase.SJsonValue;
	_sResult	: KOSTAL_AF2024_Core_Settings.T_MaxString_UTF8;
	_SP				: T_SubModuleOfProcess;
END_VAR
IF IN = 0 												THEN _getSubModule_n:= 'IN Parameter is empty';												RETURN;	END_IF
//IF Index = 0 										THEN _getSubModule_n:= 'Index is out of Range (Base = 1';							RETURN;	END_IF
IF _SubModuleListLenght = 0				THEN _getSubModule_n:= 'no content available';												RETURN;	END_IF
IF Index >= _SubModuleListLenght	THEN _getSubModule_n:= 'Index is out of Range';												RETURN;	END_IF

_J:= _JsonParser.GetArrayValueByIdx(IN,Index);

IF _J = 0	THEN _getSubModule_n:= '_getSubModule_n - no content availabe';	RETURN;	END_IF


_SP.clear();

_PARSE_STRING(_J, SUBMODUL_INFO.articleNumber, _sResult);	
_SP.articleNumber:= _sResult;

_PARSE_STRING(_J, SUBMODUL_INFO.serialNumber, _sResult);
_SP.serialNumber:= _sResult;

_PARSE_STRING(_J, SUBMODUL_INFO.timestamp, _sResult);
_SP.timeStamp:= _sResult;

_ListOfSubModules.Add_DUT(_SP, 0);

(*
IF IN = 0 THEN _getSubModules:= 'IN Parameter is empty';	RETURN;	END_IF

_sResp:= _PARSE_JSON(IN, PROCESS_INFO.processInfo, _IN);
IF _sResp <> '' THEN	_getSubModules:= _sResp;	RETURN; END_IF

_sResp:= _PARSE_ARRAY(_IN, SUBMODUL_INFO.subModules, _J);
IF _sResp <> '' THEN	_getSubModules:= _sResp;	RETURN; END_IF
IF _J = 0	THEN _getSubModules:= '_getSubModules - no content availabe';	RETURN;	END_IF

_jIterator		:= _JsonParser.ArrayBegin(_J);
_jIteratorEnd	:= _JsonParser.ArrayEnd(_J);

WHILE _jIterator <> _jIteratorEnd DO 
	
  _jElement := _JsonParser.GetArrayValue(_jIterator);
	IF _jElement = 0 THEN _getSubModules:= '_getSubModules - sub module corrupt';	RETURN;	END_IF

	_ListOfSubModules.AddObject();
	_pLoSM:= _ListOfSubModules.Get_P(_ListOfSubModules.NumberOfObjects, 0);
	
	_sResp:= _PARSE_STRING(_J, SUBMODUL_INFO.articleNumber, _sResult);
	IF _sResp <> '' THEN	_getSubModules:= _sResp;	ELSE	_pLoSM^.articleNumber:=_sResult;	END_IF

	_sResp:= _PARSE_STRING(_J, SUBMODUL_INFO.serialNumber, _sResult);
	IF _sResp <> '' THEN	_getSubModules:= _sResp;	ELSE	_pLoSM^.serialNumber:=_sResult;	END_IF

	_sResp:= _PARSE_STRING(_J, SUBMODUL_INFO.timestamp, _sResult);
	IF _sResp <> '' THEN	_getSubModules:= _sResp;	ELSE	_pLoSM^.timeStamp:=_sResult;	END_IF
	
  _jIterator := _JsonParser.NextArray(_jIterator);

END_WHILE


*)
END_METHOD

METHOD PROTECTED _getSubModuleList : KOSTAL_AF2024_Core_Settings.T_MaxString_UTF8
VAR_INPUT
	IN	: Tc3_IotBase.SJsonValue;
END_VAR

IF IN = 0 THEN _getSubModuleList:= '_getSubModuleList - IN Parameter is empty';	RETURN;	END_IF

_SubModuleListLenght:= 0;

_getSubModuleList:= _PARSE_ARRAY(IN, SUBMODUL_INFO.subModules, _JsonSubModules);

IF _getSubModuleList <> '' THEN	RETURN;	END_IF

_SubModuleListLenght:=  _JsonParser.GetArraySize(_JsonSubModules);
END_METHOD

METHOD PROTECTED _01_Ready : BOOL
VAR_INPUT
END_VAR


IF NOT 	SUPER^._01_Ready() 								THEN	

	;

ELSIF		_THIS_CALLED = E_PROCESS.idle			THEN	

	_state.clear();	
	_state.ready:= TRUE;

ELSIF		_THIS_CALLED = E_PROCESS.execute	THEN	

	_THIS_IN_PROCESS:= _THIS_CALLED;	

	_state.clear();	
	_state.busy:= TRUE;

	_selectUrl();

	_step.INC();

ELSE

	_state.clear();
	_state.fail:= TRUE;
	_state.description:= Tc2_Standard.WCONCAT("Unknown Process called:", INT_TO_WSTRING(_THIS_CALLED));
	
END_IF
END_METHOD

METHOD PROTECTED _10_getProcessInfo
VAR_INPUT
END_VAR

IF _step.toggle THEN
	;
END_IF

_sResp:= _getProcessInfo(_jsonDoc);

IF _sResp <> '' THEN
	
	_state.clear();
	_state.description:= Tc2_Standard.WCONCAT("Process Info is corrupt;", TO_WSTRING(_sResp));
	_step.set(_ADDRESS_FINISH_FAIL);

ELSE	

	_step.INC();

END_IF
END_METHOD

METHOD PROTECTED _10_getSubModule_n
VAR_INPUT
END_VAR

IF _step.toggle THEN
	;
END_IF

IF _ListOfSubModules.NumberOfMember < _SubModuleListLenght THEN

	_sResp:= _getSubModule_n(_JsonSubModules,  _ListOfSubModules.NumberOfMember);

	IF _sResp <> '' THEN
		
		_state.clear();
		_state.description:= Tc2_Standard.WCONCAT("Sub Module List is corrupt;", TO_WSTRING(_sResp));
		_step.set(_ADDRESS_FINISH_FAIL);
	
	END_IF

ELSE

	_step.INC();

END_IF


(*

_getSubModules(_JsonSubModules);

_step.INC();


//Sub modules are optional
_sResp:= _getSubModules(_jsonDoc);

IF _sResp <> '' THEN
	
	_state.clear();
	_state.description:= Tc2_Standard.CONCAT('Process Info is corrupt;', _sResp);
	_step.set(_ADDRESS_FINISH_FAIL);

ELSE	

	_step.INC();

END_IF
*)
END_METHOD

METHOD PROTECTED _10_getSubModuleList
VAR_INPUT
END_VAR

IF _step.toggle THEN
	;
END_IF

_sResp:= _getSubModuleList(_JsonProcessInfo);

IF _sResp <> '' THEN

	_state.clear();
	_state.description:= Tc2_Standard.WCONCAT("ProcessListInfo is corrupt;", TO_WSTRING(_sResp));
	
	_step.set(_ADDRESS_FINISH_FAIL);

ELSIF _SubModuleListLenght = 0 THEN
	
	_state.clear();
	_state.description:= "no SubModuleList available";

	_step.set(_ADDRESS_FINISH_FAIL);

ELSE
	
	_step.INC();

END_IF
END_METHOD

METHOD PROTECTED _10_processRead
VAR_INPUT
END_VAR

IF _step.toggle THEN

	_JsonProcessInfo:= 0;
	
	_ResponseResult.clear();
	_ResponseProcess.clear();
	_ListOfSubModules.Clear();

END_IF

_00_clientCfg();
END_METHOD

(*
| MUST EXTEND
*)
METHOD PROTECTED _selectUrl


_sUrl:= _UriGet(URL.READ_SUB_MODULES_BY_PARENT_SERIAL_NUMBER);

_UrlReplace(_sUrl, URL.PLACEHOLDER_CLIENT_NAME, _ClientName);
_UrlReplace(_sUrl, URL.PLACEHOLDER_CLIENT_PROCESS, _ClientProcess);
_UrlReplace(_sUrl, URL.PLACEHOLDER_PARENT_SERIAL_NUMBER, _SerialNumber);
END_METHOD

(*
*)
METHOD Execute : BOOL

VAR_INPUT
	SerialNumber	: KOSTAL_AF2024_Core_Settings.T_MaxString_UTF8;
END_VAR

IF _THIS_CALLED <> E_PROCESS.idle THEN Execute:= FALSE;	RETURN; END_IF

_THIS_CALLED:= E_PROCESS.execute;

IF NOT MT_Usage THEN _SerialNumber	:= SerialNumber;	end_if

_FBmain();

Execute:= _THIS_CALLED = _THIS_IN_PROCESS;
END_METHOD

PROPERTY PUBLIC ListOfSubModules : I_ListOfSubModuleOfProcess
GET

ListOfSubModules	:= _ListOfSubModules;
END_GET
END_PROPERTY

PROPERTY PUBLIC ResponseProcess : I_T_SingleProcess
GET

ResponseProcess:= _ResponseProcess;
END_GET
END_PROPERTY

PROPERTY ResponseResult : I_T_ResponseResult
GET

ResponseResult := _ResponseResult;
END_GET
END_PROPERTY

METHOD PROTECTED _FBmain
VAR_INPUT
END_VAR

SUPER^._FBmain();

CASE _step.actual OF

	0:	_01_Ready();
	//
	1:	_10_processRead();
	2:	_10_GET();
	3:	_10_GET_CTRL();
	4:	_10_GET_ResponseResult(TRUE);
	5:	_10_GET_ResponseResult_CTRL();
	6:	_10_getProcessInfo();
	7:	_10_getSubModuleList();
	8:	_10_getSubModule_n();
	9:	_10_finishPass();

	100:	_10_finishFail();
ELSE
	
	_99_stepError();
		
END_CASE
END_METHOD

END_FUNCTION_BLOCK

// 5_POU/Init/FB_Init
(*
|Extends the base WebService LC with a 
|read Process-Config with another naming
|functionality
*)
FUNCTION_BLOCK PUBLIC FB_Init EXTENDS FB_ReadProcessConfig

END_FUNCTION_BLOCK

// 5_POU/ReadProcessConfig/FB_ReadProcessConfig
(*
|Extends the base WebService LC with a 
|read config 
|functionality
================================================================================================
|if ClientProcess is not defined, the hole configuration settings for this "ClientName" is available in the response
|Otherwise only the configuration of the ClientProcess is available
*)
FUNCTION_BLOCK PUBLIC FB_ReadProcessConfig EXTENDS _FB_ReadConfig

METHOD Execute : BOOL

IF _THIS_CALLED <> E_PROCESS.idle THEN Execute:= FALSE;	RETURN; END_IF

_THIS_CALLED:= E_PROCESS.execute;

_FBmain();

Execute:= _THIS_CALLED = _THIS_IN_PROCESS;
END_METHOD

METHOD PROTECTED _selectUrl



IF _ClientProcess = '' THEN

	_sUrl:= _UriGet(URL.READ_PROC_CONF);
	_UrlReplace(_sUrl, URL.PLACEHOLDER_CLIENT_NAME, _ClientName);

ELSE

	_sUrl:= _UriGet(URL.READ_PROC_CONF_OPT_PROC);
	_UrlReplace(_sUrl, URL.PLACEHOLDER_CLIENT_NAME, _ClientName);
	_UrlReplace(_sUrl, URL.PLACEHOLDER_CLIENT_PROCESS, _ClientProcess);
	
END_IF
END_METHOD

END_FUNCTION_BLOCK

// 5_POU/ReadProcessConfig/MustBeExtended/_FB_ReadConfig
(*
|MUST EXEND
|
|Extends the base WebService LC with a 
|read configuration
|functionality
*)
FUNCTION_BLOCK ABSTRACT _FB_ReadConfig EXTENDS FB_LC

VAR

	//======================================================================================
	//Read
	//======================================================================================
	
	_ListOfConfiguration		: FB_ListOfProcessConfig;
		
	//======================================================================================
	//do not insert to _DELETE() !!!!
	_JsonProcessConfigList		: Tc3_IotBase.SJsonValue;	//do not insert to _DELETE() !!!!
	_ProcessConfigListLenght	: UDINT;									//do not insert to _DELETE() !!!!
	//======================================================================================

	
END_VAR

VAR CONSTANT
	_ADDRESS_FINISH_FAIL : INT:= 100;
END_VAR

METHOD PROTECTED _getPreviousProcess	: KOSTAL_AF2024_Core_Settings.T_MaxString_UTF8
VAR_INPUT
	jPP	: Tc3_IotBase.SJsonValue;			//PP = PreviousProcess
	PP	: I_T_PreviousProcess_Owner;	//PP = PreviousProcess
END_VAR

VAR
	_uliResult: ULINT;
	_udiResult: UDINT;
	_diResult	: DINT;
	_bResult	: BOOL;
	_sResult	: KOSTAL_AF2024_Core_Settings.T_MaxString_UTF8;
	_PP	: I_T_PreviousProcess_Owner;	//PP = PreviousProcess
END_VAR

IF jPP = 0		THEN _getPreviousProcess:= 'Json Parameter jPP is empty';	RETURN;	END_IF
IF PP = 0	THEN _getPreviousProcess:= 'Object is zero';	RETURN;	END_IF

IF NOT __QUERYINTERFACE(PP, _PP) OR_ELSE _PP = 0	THEN _getPreviousProcess:= 'Object is invalid';	RETURN;	END_IF

_PP.clear();

_sResp:= _PARSE_STRING(jPP, PROCESS_CONFIG.processName, _sResult);
IF _sResp <> '' THEN	(*ignore *) ;	ELSE	_PP.processName:= _sResult; END_IF

_sResp:= _PARSE_STRING(jPP, PROCESS_CONFIG.processStamp, _sResult);
IF _sResp <> '' THEN	(*ignore *) ;	ELSE	_PP.processStamp:= _sResult; END_IF

_sResp:= _PARSE_STRING(jPP, PROCESS_CONFIG.databaseName, _sResult);
IF _sResp <> '' THEN	(*ignore *) ;	ELSE	_PP.databaseName:= _sResult; END_IF

_sResp:= _PARSE_STRING(jPP, PROCESS_CONFIG.useOnlyTable, _sResult);
IF _sResp <> '' THEN	(*ignore *) ;	ELSE	_PP.useOnlyTable:= _sResult; END_IF

_sResp:= _PARSE_DINT(jPP, PROCESS_CONFIG.searchMode, _diResult);
IF _sResp <> '' THEN	(*ignore *) ;	ELSE	_PP.searchMode:= _diResult; END_IF

_sResp:= _PARSE_STRING(jPP, PROCESS_CONFIG.articlenumberRegex, _sResult);
IF _sResp <> '' THEN	(*ignore *) ;	ELSE	_PP.articlenumberRegex:= _sResult; END_IF

_getPreviousProcess:= _getPreviousProcesses(jPP, _PP);
END_METHOD

METHOD PROTECTED _getPreviousProcesses	: KOSTAL_AF2024_Core_Settings.T_MaxString_UTF8
VAR_INPUT
	jPP	: Tc3_IotBase.SJsonValue;			//PP = PreviousProcess
	PP	: I_T_PreviousProcess_Owner;	//PP = PreviousProcess
END_VAR

VAR
	_jPP	: Tc3_IotBase.SJsonValue;					//PP = PreviousProcesses
	_uliResult: ULINT;
	_udiResult: UDINT;
	_diResult	: DINT;
	_bResult	: BOOL;
	_sResult	: KOSTAL_AF2024_Core_Settings.T_MaxString_UTF8;
	_PP	: I_T_PreviousProcess_Owner;	//PP = PreviousProcess

	_jsonIterator			: Tc3_IotBase.SJsonIterator;
	_jsonIteratorEnd	: Tc3_IotBase.SJsonIterator;
	_jsonValue				: Tc3_IotBase.SJsonValue;
END_VAR

IF jPP = 0	THEN _getPreviousProcesses:= 'Json Parameter jPP is empty';	RETURN;	END_IF
IF PP = 0		THEN _getPreviousProcesses:= 'Object-Pointer is zero';	RETURN;	END_IF

IF NOT __QUERYINTERFACE(PP, _PP) OR_ELSE _PP = 0	THEN _getPreviousProcesses:= 'Object is invalid';	RETURN;	END_IF

_PP.PreviousProcesses_Owner.clear();

IF _PARSE_JSON(jPP, PROCESS_CONFIG.previousProcesses, _jPP) = '' THEN

	IF _jPP <> 0 THEN

		_jsonIterator := _JsonParser.MemberBegin(_jPP);
		_jsonIteratorEnd := _JsonParser.MemberEnd(_jPP);

		WHILE _jsonIterator <> _jsonIteratorEnd DO

			_jsonValue := _JsonParser.GetMemberValue(_jsonIterator);
			_PP.PreviousProcesses_Owner.addLine(_JsonParser.GetString(_jsonValue));
			
			_jsonIterator := _JsonParser.NextMember(_jsonIterator);

		END_WHILE
	
	END_IF

END_IF
END_METHOD

METHOD PROTECTED _getPreviousProcessList : KOSTAL_AF2024_Core_Settings.T_MaxString_UTF8
VAR_INPUT
	jPC	: Tc3_IotBase.SJsonValue;		//PC = ProcessConfiguration
	PC	: I_T_ProcessConfig_Owner;	//PC = ProcessConfiguration
END_VAR

VAR
	_jPrevProcessList				: Tc3_IotBase.SJsonValue;
	_PrevProcessListLenght	: UDINT;
	_jPrevProcess						: Tc3_IotBase.SJsonValue;
	_PC	: I_T_ProcessConfig_Owner;	//PC = ProcessConfiguration

	_PP	: T_PreviousProcess;	//PP = PreviousProcess
	
	_udi	: UDINT;
END_VAR

IF jPC = 0	THEN _getPreviousProcessList:= 'Json Parameter jPC is empty';	RETURN;	END_IF
IF PC = 0		THEN _getPreviousProcessList:= 'Object is zero';			RETURN;	END_IF

IF NOT __QUERYINTERFACE(PC, _PC) OR_ELSE _PC = 0	THEN _getPreviousProcessList:= 'Object is invalid';	RETURN;	END_IF

_PC.PreviousProcesses_Owner.Clear();

_sResp:= _PARSE_ARRAY(jPC, PROCESS_CONFIG.previousProcesses, _jPrevProcessList);
IF _sResp <> '' 					THEN	RETURN;	END_IF
IF _jPrevProcessList = 0	THEN	RETURN;	END_IF

_PrevProcessListLenght:=  _JsonParser.GetArraySize(_jPrevProcessList);
IF _PrevProcessListLenght = 0 THEN	RETURN;	END_IF

FOR _udi:= 1 TO _PrevProcessListLenght DO

	_jPrevProcess:= _JsonParser.GetArrayValueByIdx(_jPrevProcessList, _udi - 1);
	
	IF _jPrevProcess <> 0 THEN	
		_PP.clear();
		_getPreviousProcess(_jPrevProcess, _PP);	
		_PC.PreviousProcesses_Owner.Add_DUT(_PP, 0);
	END_IF

END_FOR
END_METHOD

(*
	| return the Process Info from List with {Index} (Base = 0)
*)
METHOD PROTECTED _getProcessConfig : KOSTAL_AF2024_Core_Settings.T_MaxString_UTF8
VAR_INPUT
	IN		: Tc3_IotBase.SJsonValue;
	Index	: UDINT;
END_VAR

VAR
	_PC	: T_ProcessConfig;	//PC = ProcessConfiguration
	_J	: Tc3_IotBase.SJsonValue;
	_uliResult: ULINT;
	_udiResult: UDINT;
	_diResult	: DINT;
	_bResult	: BOOL;
	_sResult	: KOSTAL_AF2024_Core_Settings.T_MaxString_UTF8;
	_fResp		: KOSTAL_AF2024_Core_functionResponse.T_functionResponse;
END_VAR
IF IN = 0		 													THEN _getProcessConfig:= 'IN Parameter is empty';												RETURN;	END_IF
//IF Index = 0 												THEN _getProcessInfo:= 'Index is out of Range (Base = 1';							RETURN;	END_IF
IF _ProcessConfigListLenght = 0				THEN _getProcessConfig:= 'no content available';												RETURN;	END_IF
IF Index >= _ProcessConfigListLenght 	THEN _getProcessConfig:= 'Index is out of Range';												RETURN;	END_IF

_J:= _JsonParser.GetArrayValueByIdx(IN,Index);

IF _J = 0	THEN _getProcessConfig:= '_getProcessInfo - no content availabe';	RETURN;	END_IF


//IF NOT _ListOfConfiguration.AddObject() THEN	_getProcessConfig:= 'fail during creation of ListOfConfiguration.AddObject';	RETURN; END_IF
//_PC:= _ListOfConfiguration.Get_P(_ListOfConfiguration.NumberOfObjects, _fResp);
//IF NOT _fResp.success THEN	_getProcessConfig:= _fResp.status;	RETURN; END_IF
//IF _PC = 0						THEN	_getProcessConfig:= 'fail during get Pointer to ListOfConfiguration Object';	RETURN; END_IF

_PC.clear();

_sResp:= _PARSE_STRING(_J, PROCESS_CONFIG.articlenumberRegex, _sResult);
IF _sResp <> '' THEN	_getProcessConfig:= _sResp;	ELSE	_PC.articlenumberRegex:= _sResult; END_IF

_sResp:= _PARSE_STRING(_J, PROCESS_CONFIG.serialnumberRegex, _sResult);
IF _sResp <> '' THEN	_getProcessConfig:= _sResp;	ELSE	_PC.serialnumberRegex:= _sResult;	END_IF

_sResp:= _PARSE_DINT(_J, PROCESS_CONFIG.traceID, _diResult);
IF _sResp <> '' THEN	_getProcessConfig:= _sResp;	ELSE	_PC.traceID:= _diResult;	END_IF

_sResp:= _PARSE_BOOL(_J, PROCESS_CONFIG.activeCheckFQDN, _bResult);
IF _sResp <> '' THEN	_getProcessConfig:= _sResp;	ELSE	_PC.activeCheckFQDN:= _bResult;	END_IF

_sResp:= _PARSE_STRING(_J, PROCESS_CONFIG.allowedFQDN, _sResult);
IF _sResp <> '' THEN	_getProcessConfig:= _sResp;	ELSE	_PC.allowedFQDN:= _sResult; END_IF

_getProcessConfig:= _getPreviousProcessList(_J, _PC);

IF _getProcessConfig = '' THEN	_ListOfConfiguration.Add_DUT(_PC, 0);	END_IF
END_METHOD

METHOD PROTECTED _getProcessConfigList : KOSTAL_AF2024_Core_Settings.T_MaxString_UTF8
VAR_INPUT
	IN	: Tc3_IotBase.SJsonValue;
END_VAR

IF IN = 0 THEN _getProcessConfigList:= '_getProcessConfigList - IN Parameter is empty';	RETURN;	END_IF

_ProcessConfigListLenght:= 0;

_getProcessConfigList:= _PARSE_ARRAY(IN, PROCESS_CONFIG.processConfiguration, _JsonProcessConfigList);

IF _getProcessConfigList <> '' THEN	RETURN;	END_IF

_ProcessConfigListLenght:=  _JsonParser.GetArraySize(_JsonProcessConfigList);
END_METHOD

METHOD PROTECTED _01_Ready : BOOL
VAR_INPUT
END_VAR


IF NOT 	SUPER^._01_Ready() 								THEN	

	;

ELSIF		_THIS_CALLED = E_PROCESS.idle			THEN	

	_state.clear();	
	_state.ready:= TRUE;

ELSIF		_THIS_CALLED = E_PROCESS.execute	THEN	

	_THIS_IN_PROCESS:= _THIS_CALLED;	

	_state.clear();	
	_state.busy:= TRUE;

	_selectUrl();

	_step.INC();

ELSE

	_state.clear();
	_state.fail:= TRUE;
	_state.description:= Tc2_Standard.WCONCAT("Unknown Process called:", INT_TO_WSTRING(_THIS_CALLED));
	
END_IF
END_METHOD

METHOD PROTECTED _10_getProcessConfig_n

VAR
	_c	: KOSTAL_AF2024_Core_StringTools.FB_Concat;
END_VAR

IF _step.toggle THEN
	;
END_IF

IF _ListOfConfiguration.NumberOfMember < _ProcessConfigListLenght THEN

	_sResp:= _getProcessConfig(_JsonProcessConfigList,  _ListOfConfiguration.NumberOfMember);

	IF _sResp <> '' THEN
	
		_state.clear();

		_c.clear();
		_c.addContent("Process Info ");
		_c.addContent(UDINT_TO_WSTRING(_ListOfConfiguration.NumberOfMember));
		_c.addContent(" is corrupt;");
		_c.addContent(TO_WSTRING(_sResp));
		_state.description:= _c.getResult();
		_c.clear();

		_step.set(_ADDRESS_FINISH_FAIL);

	END_IF
	
ELSE

	_step.INC();

END_IF
END_METHOD

METHOD PROTECTED _10_getProcessConfigList
VAR_INPUT
END_VAR

IF _step.toggle THEN
	;
END_IF

_sResp:= _getProcessConfigList(_jsonDoc);

IF _sResp <> '' THEN

	_state.clear();
	_state.description:= Tc2_Standard.WCONCAT("ProcessConfigList is corrupt;", TO_WSTRING(_sResp));
	
	_step.set(_ADDRESS_FINISH_FAIL);

ELSIF _ProcessConfigListLenght = 0 THEN
	
	_state.clear();
	_state.description:= "no ProcessListInfo available";

	_step.set(_ADDRESS_FINISH_FAIL);

ELSE
	
	_step.INC();

END_IF
END_METHOD

METHOD PROTECTED _10_processRead
VAR_INPUT
END_VAR

IF _step.toggle THEN

	_JsonProcessConfigList:= 0;

	_ResponseResult.clear();

	_ListOfConfiguration.Clear();

END_IF

_00_clientCfg();
END_METHOD

(*
| MUST EXTEND
*)
METHOD PROTECTED _selectUrl
END_METHOD

METHOD PUBLIC GetProcessConfig : I_T_ProcessConfig
VAR_INPUT
	ListNumber	: UDINT;
END_VAR

GetProcessConfig:= _ListOfConfiguration.Get_I(ListNumber, 0, 0);
END_METHOD

PROPERTY PUBLIC NumberOfProcessConfig : UDINT
GET

NumberOfProcessConfig:= _ListOfConfiguration.NumberOfMember;
END_GET
END_PROPERTY

PROPERTY ResponseResult : I_T_ResponseResult
GET

ResponseResult := _ResponseResult;
END_GET
END_PROPERTY

METHOD PROTECTED _FBmain
VAR_INPUT
END_VAR

SUPER^._FBmain();

CASE _step.actual OF

	0:	_01_Ready();
	//
	1:	_10_processRead();
	2:	_10_GET();
	3:	_10_GET_CTRL();
	4:	_10_GET_ResponseResult(TRUE);
	5:	_10_GET_ResponseResult_CTRL();
	6:	_10_getProcessConfigList();
	7:	_10_getProcessConfig_n();
	8:	_10_finishPass();

	100:	_10_finishFail();
ELSE
	
	_99_stepError();
		
END_CASE
END_METHOD

END_FUNCTION_BLOCK

// 5_POU/ReadApiVersion/MustBeExtended/_FB_ReadApiVersion
(*
|MUST EXEND
|
|Extends the base WebService LC with a 
|read
|and a 
|read previous Stamp 
|functionality
*)
FUNCTION_BLOCK ABSTRACT _FB_ReadApiVersion EXTENDS FB_LC

VAR
	_apiVersion	: KOSTAL_AF2024_Core_Settings.T_MaxString_UTF8;
END_VAR

VAR CONSTANT
	_ADDRESS_FINISH_FAIL : INT:= 100;
END_VAR

METHOD PROTECTED _getApiVersion : KOSTAL_AF2024_Core_Settings.T_MaxString_UTF8
VAR_INPUT
	IN	: Tc3_IotBase.SJsonValue;
END_VAR

VAR
	_sResult: KOSTAL_AF2024_Core_Settings.T_MaxString_UTF8;
END_VAR

_apiVersion:= '';

IF IN = 0 THEN _getApiVersion:= '_getApiVersion - IN Parameter is empty';	RETURN;	END_IF

_sResp:= _PARSE_STRING(IN, API_VERSION.apiVersion, _sResult);

IF _sResp <> '' THEN	_getApiVersion:= _sResp;	ELSE	_apiVersion:= _sResult;	END_IF
END_METHOD

METHOD PROTECTED _01_Ready : BOOL
VAR_INPUT
END_VAR


IF NOT 	SUPER^._01_Ready() 								THEN	

	;

ELSIF		_THIS_CALLED = E_PROCESS.idle			THEN	

	_state.clear();	
	_state.ready:= TRUE;

ELSIF		_THIS_CALLED = E_PROCESS.execute	THEN	

	_THIS_IN_PROCESS:= _THIS_CALLED;	

	_state.clear();	
	_state.busy:= TRUE;

	_selectUrl();

	_step.INC();

ELSE

	_state.clear();
	_state.fail:= TRUE;
	_state.description:= Tc2_Standard.WCONCAT("Unknown Process called:", INT_TO_WSTRING(_THIS_CALLED));
	
END_IF
END_METHOD

METHOD PROTECTED _10_getapiVersion
VAR_INPUT
END_VAR

IF _step.toggle THEN
	;
END_IF

_sResp:= _getApiVersion(_jsonDoc);

IF _sResp <> '' THEN

	_state.clear();
	_state.description:= Tc2_Standard.WCONCAT("ProcessListInfo is corrupt;", TO_WSTRING(_sResp));
	
	_step.set(_ADDRESS_FINISH_FAIL);

ELSE
	
	_step.INC();

END_IF
END_METHOD

METHOD PROTECTED _10_processRead
VAR_INPUT
END_VAR

IF _step.toggle THEN

	_ResponseResult.clear();

END_IF

_00_clientCfg();
END_METHOD

(*
| MUST EXTEND
*)
METHOD PROTECTED _selectUrl
END_METHOD

PROPERTY PUBLIC apiVersion : KOSTAL_AF2024_Core_Settings.T_MaxString_UTF8
GET

apiVersion:= _apiVersion;
END_GET
END_PROPERTY

PROPERTY ResponseResult : I_T_ResponseResult
GET

ResponseResult := _ResponseResult;
END_GET
END_PROPERTY

METHOD PROTECTED _FBmain
VAR_INPUT
END_VAR

SUPER^._FBmain();

CASE _step.actual OF

	0:	_01_Ready();
	//
	1:	_10_processRead();
	2:	_10_GET();
	3:	_10_GET_CTRL();
	4:	_10_GET_ResponseResult(TRUE);
	5:	_10_GET_ResponseResult_CTRL();
	6:	_10_getapiVersion();
	7:	_10_finishPass();

	100:	_10_finishFail();
ELSE
	
	_99_stepError();
		
END_CASE
END_METHOD

END_FUNCTION_BLOCK

// 5_POU/ReadApiVersion/FB_ReadApiVersion
(*
|Extends the base WebService LC with a 
|read
|and a 
|read previous Stamp 
|functionality
*)
FUNCTION_BLOCK PUBLIC FB_ReadApiVersion EXTENDS _FB_ReadApiVersion

METHOD Execute : BOOL

IF _THIS_CALLED <> E_PROCESS.idle THEN Execute:= FALSE;	RETURN; END_IF

_THIS_CALLED:= E_PROCESS.execute;

_FBmain();

Execute:= _THIS_CALLED = _THIS_IN_PROCESS;
END_METHOD

METHOD PROTECTED _selectUrl


_sUrl:= _UriGet(URL.READ_API_VERSION);
END_METHOD

END_FUNCTION_BLOCK

// 5_POU/ReadProcess/MustBeExtended/_FB_ReadProcess
(*
|MUST EXEND
|
|Extends the base WebService LC with a 
|read
|and a 
|read previous Stamp 
|functionality
*)
FUNCTION_BLOCK ABSTRACT _FB_ReadProcess EXTENDS FB_LC

VAR

	//======================================================================================
	//Read
	//======================================================================================
	
	_ListOfSingleProcess		: FB_ListOfSingleProcess;
		
	//======================================================================================
	//do not insert to _DELETE() !!!!
	_JsonProcessInfoList: Tc3_IotBase.SJsonValue;	//do not insert to _DELETE() !!!!
	_ProcessInfoListLenght	: UDINT;								//do not insert to _DELETE() !!!!
	//======================================================================================

	
END_VAR

VAR CONSTANT
	_ADDRESS_FINISH_FAIL : INT:= 100;
END_VAR

(*
	| return the Process Info from List with {Index} (Base = 0)
*)
METHOD PROTECTED _getProcessInfo : KOSTAL_AF2024_Core_Settings.T_MaxString_UTF8
VAR_INPUT
	IN		: Tc3_IotBase.SJsonValue;
	Index	: UDINT;
END_VAR

VAR
	_SP	: T_SingleProcess;	//SP = SingleProcess
	_J	: Tc3_IotBase.SJsonValue;
	_uliResult: ULINT;
	_udiResult: UDINT;
	_diResult	: DINT;
	_bResult	: BOOL;
	_sResult	: KOSTAL_AF2024_Core_Settings.T_MaxString_UTF8;
END_VAR

IF IN = 0 												THEN _getProcessInfo:= 'IN Parameter is empty';							RETURN;	END_IF
//IF Index = 0 											THEN _getProcessInfo:= 'Index is out of Range (Base = 1';	RETURN;	END_IF
IF _ProcessInfoListLenght = 0			THEN _getProcessInfo:= 'no content available';							RETURN;	END_IF
IF Index >= _ProcessInfoListLenght THEN _getProcessInfo:= 'Index is out of Range';						RETURN;	END_IF

_J:= _JsonParser.GetArrayValueByIdx(IN,Index);

IF _J = 0	THEN _getProcessInfo:= '_getProcessInfo - no content availabe';	RETURN;	END_IF

_SP.clear();

_sResp:= _PARSE_ULINT(_J, PROCESS_INFO.id, _uliResult);
IF _sResp <> '' THEN	_getProcessInfo:= _sResp;	ELSE	_SP.id:= _uliResult; END_IF

_sResp:= _PARSE_STRING(_J, PROCESS_INFO.serialNumber, _sResult);
IF _sResp <> '' THEN	_getProcessInfo:= _sResp;	ELSE	_SP.serialNumber:= _sResult;	END_IF

_sResp:= _PARSE_STRING(_J, PROCESS_INFO.articleNumber, _sResult);
IF _sResp <> '' THEN	_getProcessInfo:= _sResp;	ELSE	_SP.articleNumber:= _sResult;	END_IF

_sResp:= _PARSE_STRING(_J, PROCESS_INFO.timeStamp, _sResult);
IF _sResp <> '' THEN	_getProcessInfo:= _sResp;	ELSE	_SP.timeStamp:= _sResult;	END_IF

_sResp:= _PARSE_DINT(_J, PROCESS_INFO.traceId, _diResult);
IF _sResp <> '' THEN	_getProcessInfo:= _sResp;	ELSE	_SP.traceId:= _diResult; END_IF

_sResp:= _PARSE_STRING(_J, PROCESS_INFO.process, _sResult);
IF _sResp <> '' THEN	_getProcessInfo:= _sResp;	ELSE	_SP.process:= _sResult;	END_IF

_sResp:= _PARSE_BOOL(_J, PROCESS_INFO.result, _bResult);
IF _sResp <> '' THEN	_getProcessInfo:= _sResp;	ELSE	_SP.result:= _bResult;	END_IF

_sResp:= _PARSE_STRING(_J, PROCESS_INFO.optionalString_1, _sResult);
IF _sResp <> '' THEN	_getProcessInfo:= _sResp;	ELSE	_SP.OptionalStrings_Owner.set(1, _sResult);	END_IF

_sResp:= _PARSE_STRING(_J, PROCESS_INFO.optionalString_2, _sResult);
IF _sResp <> '' THEN	_getProcessInfo:= _sResp;	ELSE	_SP.OptionalStrings_Owner.set(2, _sResult);	END_IF

_sResp:= _PARSE_STRING(_J, PROCESS_INFO.optionalString_3, _sResult);
IF _sResp <> '' THEN	_getProcessInfo:= _sResp;	ELSE	_SP.OptionalStrings_Owner.set(3, _sResult);	END_IF

_sResp:= _PARSE_STRING(_J, PROCESS_INFO.optionalString_4, _sResult);
IF _sResp <> '' THEN	_getProcessInfo:= _sResp;	ELSE	_SP.OptionalStrings_Owner.set(4, _sResult);	END_IF

_sResp:= _PARSE_BOOL(_J, PROCESS_INFO.optionalFlag_1, _bResult);
IF _sResp <> '' THEN	_getProcessInfo:= _sResp;	ELSE	_SP.OptionalFlags_Owner.set(1, (_bResult <> 0));	END_IF

_sResp:= _PARSE_BOOL(_J, PROCESS_INFO.optionalFlag_2, _bResult);
IF _sResp <> '' THEN	_getProcessInfo:= _sResp;	ELSE	_SP.OptionalFlags_Owner.set(2, (_bResult <> 0));	END_IF

_sResp:= _PARSE_BOOL(_J, PROCESS_INFO.optionalFlag_3, _bResult);
IF _sResp <> '' THEN	_getProcessInfo:= _sResp;	ELSE	_SP.OptionalFlags_Owner.set(3, (_bResult <> 0));	END_IF

_sResp:= _PARSE_BOOL(_J, PROCESS_INFO.optionalFlag_4, _bResult);
IF _sResp <> '' THEN	_getProcessInfo:= _sResp;	ELSE	_SP.OptionalFlags_Owner.set(4, (_bResult <> 0));	END_IF

_sResp:= _PARSE_BOOL(_J, PROCESS_INFO.optionalFlag_5, _bResult);
IF _sResp <> '' THEN	_getProcessInfo:= _sResp;	ELSE	_SP.OptionalFlags_Owner.set(5, (_bResult <> 0));	END_IF

_sResp:= _PARSE_BOOL(_J, PROCESS_INFO.optionalFlag_6, _bResult);
IF _sResp <> '' THEN	_getProcessInfo:= _sResp;	ELSE	_SP.OptionalFlags_Owner.set(6, (_bResult <> 0));	END_IF

_sResp:= _PARSE_BOOL(_J, PROCESS_INFO.optionalFlag_7, _bResult);
IF _sResp <> '' THEN	_getProcessInfo:= _sResp;	ELSE	_SP.OptionalFlags_Owner.set(7, (_bResult <> 0));	END_IF

_sResp:= _PARSE_BOOL(_J, PROCESS_INFO.optionalFlag_8, _bResult);
IF _sResp <> '' THEN	_getProcessInfo:= _sResp;	ELSE	_SP.OptionalFlags_Owner.set(8, (_bResult <> 0));	END_IF

_ListOfSingleProcess.Add_DUT(_SP, 0);
END_METHOD

METHOD PROTECTED _getProcessInfoList : KOSTAL_AF2024_Core_Settings.T_MaxString_UTF8
VAR_INPUT
	IN	: Tc3_IotBase.SJsonValue;
END_VAR

IF IN = 0 THEN _getProcessInfoList:= '_getProcessInfoList - IN Parameter is empty';	RETURN;	END_IF

_ProcessInfoListLenght:= 0;

_getProcessInfoList:= _PARSE_ARRAY(IN, PROCESS_INFO.processInfoList, _JsonProcessInfoList);

IF _getProcessInfoList <> '' THEN	RETURN;	END_IF

_ProcessInfoListLenght:=  _JsonParser.GetArraySize(_JsonProcessInfoList);
END_METHOD

METHOD PROTECTED _01_Ready : BOOL
VAR_INPUT
END_VAR


IF NOT 	SUPER^._01_Ready() 								THEN	

	;

ELSIF		_THIS_CALLED = E_PROCESS.idle			THEN	

	_state.clear();	
	_state.ready:= TRUE;

ELSIF		_THIS_CALLED = E_PROCESS.execute	THEN	

	_THIS_IN_PROCESS:= _THIS_CALLED;	

	_state.clear();	
	_state.busy:= TRUE;

	_selectUrl();

	_step.INC();

ELSE

	_state.clear();
	_state.fail:= TRUE;
	_state.description:= Tc2_Standard.WCONCAT("Unknown Process called:", INT_TO_WSTRING(_THIS_CALLED));
	
END_IF
END_METHOD

METHOD PROTECTED _10_getProcessInfo_n
VAR
	_c	: KOSTAL_AF2024_Core_StringTools.FB_Concat;
END_VAR

IF _step.toggle THEN
	;
END_IF

IF _ListOfSingleProcess.NumberOfMember < _ProcessInfoListLenght THEN

	_sResp:= _getProcessInfo(_JsonProcessInfoList,  _ListOfSingleProcess.NumberOfMember);

	IF _sResp <> '' THEN
	
		_state.clear();

		_c.clear();
		_c.addContent("Process Info ");
		_c.addContent(UDINT_TO_WSTRING(_ListOfSingleProcess.NumberOfMember));
		_c.addContent(" is corrupt;");
		_c.addContent(TO_WSTRING(_sResp));
		_state.description:= _c.getResult();
		_c.clear();

		_step.set(_ADDRESS_FINISH_FAIL);

	END_IF
	
ELSE

	_step.INC();

END_IF
END_METHOD

METHOD PROTECTED _10_getProcessInfoList
VAR_INPUT
END_VAR

IF _step.toggle THEN
	;
END_IF

_sResp:= _getProcessInfoList(_jsonDoc);

IF _sResp <> '' THEN

	_state.clear();
	_state.description:= Tc2_Standard.WCONCAT("ProcessListInfo is corrupt;", TO_WSTRING(_sResp));
	
	_step.set(_ADDRESS_FINISH_FAIL);

ELSIF _ProcessInfoListLenght = 0 THEN
	
	_state.clear();
	_state.description:= "no ProcessListInfo available";

	_step.set(_ADDRESS_FINISH_FAIL);

ELSE
	
	_step.INC();

END_IF
END_METHOD

METHOD PROTECTED _10_processRead
VAR_INPUT
END_VAR

IF _step.toggle THEN

	_JsonProcessInfoList:= 0;

	_ResponseResult.clear();

	_ListOfSingleProcess.Clear();

END_IF

_00_clientCfg();
END_METHOD

(*
| MUST EXTEND
*)
METHOD PROTECTED _selectUrl
END_METHOD

METHOD PUBLIC GetSingleProcess : I_T_SingleProcess
VAR_INPUT
	ListNumber	: UDINT;
END_VAR

GetSingleProcess:= _ListOfSingleProcess.Get_I(ListNumber, 0, 0);
END_METHOD

PROPERTY PUBLIC NumberOfSingleProcess : UDINT
GET

NumberOfSingleProcess:= _ListOfSingleProcess.NumberOfMember;
END_GET
END_PROPERTY

(*
	| returns the Quantitiy of Recors in LC-Response
*)
PROPERTY ProcessInfoListLenght : UDINT
GET

ProcessInfoListLenght:= _ProcessInfoListLenght;
END_GET
END_PROPERTY

PROPERTY ResponseResult : I_T_ResponseResult
GET

ResponseResult := _ResponseResult;
END_GET
END_PROPERTY

METHOD PROTECTED _FBmain
VAR_INPUT
END_VAR

SUPER^._FBmain();

CASE _step.actual OF

	0:	_01_Ready();
	//
	1:	_10_processRead();
	2:	_10_GET();
	3:	_10_GET_CTRL();
	4:	_10_GET_ResponseResult(TRUE);
	5:	_10_GET_ResponseResult_CTRL();
	6:	_10_getProcessInfoList();
	7:	_10_getProcessInfo_n();
	8:	_10_finishPass();

	100:	_10_finishFail();
ELSE
	
	_99_stepError();
		
END_CASE
END_METHOD

END_FUNCTION_BLOCK

// 5_POU/ReadProcess/FB_ReadPreviousProcess_SN
(*
|Extends the base WebService LC with a 
|read
|and a 
|read previous Stamp 
|functionality
*)
FUNCTION_BLOCK PUBLIC FB_ReadPreviousProcess_SN EXTENDS _FB_ReadProcess

VAR
	_SerialNumber			: KOSTAL_AF2024_Core_Settings.T_MaxString_UTF8;
	_OptionalProcess	: KOSTAL_AF2024_Core_Settings.T_MaxString_UTF8;
END_VAR

METHOD Execute : BOOL

VAR_INPUT
	SerialNumber		: KOSTAL_AF2024_Core_Settings.T_MaxString_UTF8;
END_VAR

IF _THIS_CALLED <> E_PROCESS.idle THEN Execute:= FALSE;	RETURN; END_IF

_THIS_CALLED:= E_PROCESS.execute;

IF NOT MT_Usage THEN _SerialNumber	:= SerialNumber;	END_IF

_FBmain();

Execute:= _THIS_CALLED = _THIS_IN_PROCESS;
END_METHOD

METHOD PROTECTED _selectUrl


_sUrl:= _UriGet(URL.READ_PREV_PROC_SERNO);

_UrlReplace(_sUrl, URL.PLACEHOLDER_CLIENT_NAME, _ClientName);
_UrlReplace(_sUrl, URL.PLACEHOLDER_CLIENT_PROCESS, _ClientProcess);
_UrlReplace(_sUrl, URL.PLACEHOLDER_SERIALNUMBER, _SerialNumber);
END_METHOD

END_FUNCTION_BLOCK

// 5_POU/ReadProcess/FB_ReadPreviousProcess_SN_ART
(*
|Extends the base WebService LC with a 
|read
|and a 
|read previous Stamp 
|functionality
*)
FUNCTION_BLOCK PUBLIC FB_ReadPreviousProcess_SN_ART EXTENDS _FB_ReadProcess

VAR
	_SerialNumber			: KOSTAL_AF2024_Core_Settings.T_MaxString_UTF8;
	_ArticleNumber		: KOSTAL_AF2024_Core_Settings.T_MaxString_UTF8;
END_VAR

(*
|Process is an optional parameter.
|set to '' (empty string) if not used
*)
METHOD Execute : BOOL

VAR_INPUT
	SerialNumber		: KOSTAL_AF2024_Core_Settings.T_MaxString_UTF8;
	ArticleNumber		: KOSTAL_AF2024_Core_Settings.T_MaxString_UTF8;
END_VAR

IF _THIS_CALLED <> E_PROCESS.idle THEN Execute:= FALSE;	RETURN; END_IF

_THIS_CALLED:= E_PROCESS.execute;

IF NOT MT_Usage THEN 
	_SerialNumber			:= SerialNumber;
	_ArticleNumber		:= ArticleNumber;
END_IF

_FBmain();

Execute:= _THIS_CALLED = _THIS_IN_PROCESS;
END_METHOD

METHOD PROTECTED _selectUrl


_sUrl:= _UriGet(URL.READ_PREV_PROC_SERNO_ARTNO);

_UrlReplace(_sUrl, URL.PLACEHOLDER_CLIENT_NAME, _ClientName);
_UrlReplace(_sUrl, URL.PLACEHOLDER_CLIENT_PROCESS, _ClientProcess);
_UrlReplace(_sUrl, URL.PLACEHOLDER_SERIALNUMBER, _SerialNumber);
_UrlReplace(_sUrl, URL.PLACEHOLDER_ARTICLENUMBER, _ArticleNumber);
END_METHOD

END_FUNCTION_BLOCK

// 5_POU/ReadProcess/FB_ReadProcess_ID
(*
|Extends the base WebService LC with a 
|read
|and a 
|read previous Stamp 
|functionality
*)
FUNCTION_BLOCK PUBLIC FB_ReadProcess_ID EXTENDS _FB_ReadProcess

VAR
	_Record_ID	: KOSTAL_AF2024_Core_Settings.T_MaxString_UTF8;
END_VAR

METHOD Execute : BOOL

VAR_INPUT
	Record_ID	: KOSTAL_AF2024_Core_Settings.T_MaxString_UTF8;
END_VAR

IF _THIS_CALLED <> E_PROCESS.idle THEN Execute:= FALSE;	RETURN; END_IF

_THIS_CALLED:= E_PROCESS.execute;

IF NOT MT_Usage THEN _Record_ID	:= Record_ID;	END_IF

_FBmain();

Execute:= _THIS_CALLED = _THIS_IN_PROCESS;
END_METHOD

METHOD PROTECTED _selectUrl


_sUrl:= _UriGet(URL.READ_PROC_RECORD_ID);

_UrlReplace(_sUrl, URL.PLACEHOLDER_CLIENT_NAME, _ClientName);
_UrlReplace(_sUrl, URL.PLACEHOLDER_CLIENT_PROCESS, _ClientProcess);
_UrlReplace(_sUrl, URL.PLACEHOLDER_RECORD_ID, _Record_ID);
END_METHOD

END_FUNCTION_BLOCK

// 5_POU/ReadProcess/FB_ReadProcess_SN
(*
|Extends the base WebService LC with a 
|read
|and a 
|read previous Stamp 
|functionality
*)
FUNCTION_BLOCK PUBLIC FB_ReadProcess_SN EXTENDS _FB_ReadProcess

VAR
	_SerialNumber			: KOSTAL_AF2024_Core_Settings.T_MaxString_UTF8;
	_OptionalProcess	: KOSTAL_AF2024_Core_Settings.T_MaxString_UTF8;
END_VAR

(*
|Process is an optional parameter.
|set to '' (empty string) if not used
*)
METHOD Execute : BOOL

VAR_INPUT
	SerialNumber		: KOSTAL_AF2024_Core_Settings.T_MaxString_UTF8;
	OptionalProcess	: KOSTAL_AF2024_Core_Settings.T_MaxString_UTF8:= ''; //OPTIONAL
END_VAR

IF _THIS_CALLED <> E_PROCESS.idle THEN Execute:= FALSE;	RETURN; END_IF

_THIS_CALLED:= E_PROCESS.execute;

IF NOT MT_Usage THEN 
	_SerialNumber			:= SerialNumber;
	_OptionalProcess	:= OptionalProcess;
END_IF

_FBmain();

Execute:= _THIS_CALLED = _THIS_IN_PROCESS;
END_METHOD

METHOD PROTECTED _selectUrl

IF _OptionalProcess = '' THEN
	_sUrl:= _UriGet(URL.READ_PROC_SERNO);
ELSE
	_sUrl:= _UriGet(URL.READ_PROCESS_SERNO_OPT_PROC);
	_UrlReplace(_sUrl, URL.PLACEHOLDER_OPTIONAL_PROCESS, _OptionalProcess);
END_IF

_UrlReplace(_sUrl, URL.PLACEHOLDER_CLIENT_NAME, _ClientName);
_UrlReplace(_sUrl, URL.PLACEHOLDER_CLIENT_PROCESS, _ClientProcess);
_UrlReplace(_sUrl, URL.PLACEHOLDER_SERIALNUMBER, _SerialNumber);
END_METHOD

END_FUNCTION_BLOCK

// 5_POU/ReadProcess/FB_ReadProcess_SN_ART
(*
|Extends the base WebService LC with a 
|read
|and a 
|read previous Stamp 
|functionality
*)
FUNCTION_BLOCK PUBLIC FB_ReadProcess_SN_ART EXTENDS _FB_ReadProcess

VAR
	_SerialNumber			: KOSTAL_AF2024_Core_Settings.T_MaxString_UTF8;
	_ArticleNumber		: KOSTAL_AF2024_Core_Settings.T_MaxString_UTF8;
	_OptionalProcess	: KOSTAL_AF2024_Core_Settings.T_MaxString_UTF8;
END_VAR

(*
|Process is an optional parameter.
|set to '' (empty string) if not used
*)
METHOD Execute : BOOL

VAR_INPUT
	SerialNumber		: KOSTAL_AF2024_Core_Settings.T_MaxString_UTF8;
	ArticleNumber		: KOSTAL_AF2024_Core_Settings.T_MaxString_UTF8;
	OptionalProcess	: KOSTAL_AF2024_Core_Settings.T_MaxString_UTF8:= ''; //OPTIONAL
END_VAR

IF _THIS_CALLED <> E_PROCESS.idle THEN Execute:= FALSE;	RETURN; END_IF

_THIS_CALLED:= E_PROCESS.execute;

IF NOT MT_Usage THEN 
	_SerialNumber			:= SerialNumber;
	_ArticleNumber		:= ArticleNumber;
	_OptionalProcess	:= OptionalProcess;
END_IF

_FBmain();

Execute:= _THIS_CALLED = _THIS_IN_PROCESS;
END_METHOD

METHOD PROTECTED _selectUrl

IF _OptionalProcess = '' THEN

	_sUrl:= _UriGet(URL.READ_PROC_SERNO_ARTNO);

ELSE
	
	_sUrl:= _UriGet(URL.READ_PROC_SERNO_ARTNO_OPT_PROC);

	_UrlReplace(_sUrl, URL.PLACEHOLDER_OPTIONAL_PROCESS, _OptionalProcess);

END_IF

_UrlReplace(_sUrl, URL.PLACEHOLDER_CLIENT_NAME, _ClientName);
_UrlReplace(_sUrl, URL.PLACEHOLDER_CLIENT_PROCESS, _ClientProcess);
_UrlReplace(_sUrl, URL.PLACEHOLDER_SERIALNUMBER, _SerialNumber);
_UrlReplace(_sUrl, URL.PLACEHOLDER_ARTICLENUMBER, _ArticleNumber);
END_METHOD

END_FUNCTION_BLOCK

// 5_POU/WriteProcess/MustBeExtended/_FB_WriteProcess
(*
|MUST EXEND
|
|Extends the base WebService LC with a 
|write
|functionality
*)
FUNCTION_BLOCK ABSTRACT _FB_WriteProcess EXTENDS FB_LC

VAR

	//======================================================================================
	//Parameter
	//======================================================================================
	
	_WriteDataDto	: T_WriteCurrentStampDataDto;
	

	//======================================================================================
	//Response
	//======================================================================================

	_ResponseProcess: T_SingleProcess;

END_VAR

VAR CONSTANT
	_ADDRESS_FINISH_FAIL : INT:= 100;
END_VAR

